(* PLC project HomeAutomation.ecp, WAGO e!COCKPIT e!COCKPIT *)
(* stored: creationDateTime 2022-11-14T18:30:35.868664, modificationDateTime 2022-11-14T18:29:50.9667677 *)

TYPE COVER_STATES : (Idle, Auto, Manual, Prio_up, Prio_dn, Calibrate_up, Calibrate_dn);
END_TYPE

TYPE MQTT_MESSAGE : STRUCT
  Payload : STRING(128);
  Topic : STRING(128);
  Qos : MQTT.QoS;
  MqttRetain : BOOL;
END_STRUCT;
END_TYPE

TYPE RS485_EASTRON_SDM_Devices : (SDM120, SDM220, SDM630);
END_TYPE

TYPE RS485_RtuQuery : STRUCT
  DeviceId : BYTE;
  FunctionCode : BYTE;
  ReadAddress : UINT;
  ReadQuantity : UINT;
END_STRUCT;
END_TYPE

TYPE VIRTUAL_MODES : (Input, Output);
END_TYPE

INTERFACE RS485Device
METHOD RequestBusTime : BOOL
END_METHOD
METHOD GetRtuQuery : RS485_RtuQuery
END_METHOD
METHOD ProcessDataArray
  VAR_INPUT
    Error : POINTER TO BOOL;
    Data : POINTER TO ARRAY[0..124] OF WORD;
  END_VAR
END_METHOD
END_INTERFACE

FUNCTION_BLOCK _RMP_B
  VAR_INPUT
    DIR : BOOL;  (* true = up *)
    E : BOOL := TRUE;
    TR : TIME;
  END_VAR
  VAR_IN_OUT
    RMP : BYTE;
  END_VAR
  VAR
    tx : TIME;
    tl : TIME;
    tn : TIME;
    init : BOOL;
    last_dir : BOOL;
    start : BYTE;
  END_VAR

            (* read system timer *)
tx := DWORD_TO_TIME(OSCAT_BASIC.T_PLC_MS());

IF E AND init AND (dir = last_dir) AND (RMP <> SEL(DIR, 0, 255)) AND TR = tn THEN
	RMP := OSCAT_BASIC.FRMP_B(start, DIR, tx - tl, TR);
ELSE
	init := TRUE;
	tl := tx;
	tn := tr;
	start := RMP;
END_IF;
last_dir := dir;



(* revison history
hm	22. oct. 2008	rev 1.0
	original version

hm	20. nov. 2008	rev 1.1
	set default for E to be TRUE
	added init

hm	19. nov. 2011	rev 1.2
	new code
*)
          

METHOD SetRMP
  VAR_INPUT
    RMP : BYTE;
  END_VAR
                  (*THIS^.RMP:=RMP;*)
THIS^.Start:=RMP;
                
END_METHOD
END_FUNCTION_BLOCK

FUNCTION_BLOCK BLIND_ACTUATOR
  VAR_INPUT
    UP : BOOL;
    DN : BOOL;
    S_IN : BYTE;
    T_UD : TIME := TIME#10s0ms;
    T_ANGLE : TIME := TIME#3s0ms;
    {attribute 'input_constant'}
    T_LOCKOUT : TIME := TIME#100ms;
  END_VAR
  VAR_OUTPUT
    POS : BYTE;
    ANG : BYTE;
    QU : BOOL;
    QD : BOOL;
    STATUS : BYTE;
  END_VAR
  VAR
    position : RMP_B;
    angle : RMP_B;
    lock : OSCAT_BASIC.INTERLOCK;
  END_VAR

            (* make sure only one motor is active at a given time *)
lock(i1 := UP, I2 := DN, TL := T_lockout);

(* ramp up or down to simulate the angle position of the blind slats *)
angle(e := lock.Q1 OR lock.Q2, UP := lock.Q1, PT := T_Angle);
position(e := lock.Q1 AND angle.high OR lock.Q2 AND angle.low, up := lock.Q1, PT := T_UD);

(* set the outputs *)
pos := position.Out;
ang := angle.Out;

(* set the outputs *)
QU := lock.Q1;
QD := lock.Q2;

(* set the status output *)
IF UP AND DN THEN
	 status := 1;			(* error up and down together are not allowed *)
ELSIF UP THEN
	status := 121;
ELSIF DN THEN
	status := 122;
ELSE
	status := S_IN;
END_IF;


(* revision history
hm	29. sep 2007	rev 1.0
	original release

hm	6. oct 2007	rev 1.1
	rearanged outputs

hm	18. oct. 2008	rev 1.2
	changed calls for rmp_B because of change in RMP_B

hm	27. jul. 2009	rev 1.3
	changes status to be 12X

ae	08. mar. 2010 rev 1.4	
	at aPosition

*)
          

METHOD SetPOS
  VAR_INPUT
    POS : BYTE;
  END_VAR
                  THIS^.POS:=POS;
THIS^.position.SetRMP(POS);
                
END_METHOD
END_FUNCTION_BLOCK

FUNCTION CALC_COVER_STATE : COVER_STATES
  VAR_INPUT
    UP : BOOL;
    DN : BOOL;
    PRIO_LOCK : BOOL;
    PRIO_UP : BOOL;
    PRIO_DN : BOOL;
    PI : BYTE;
    POS : BYTE;
    MqttRequestAuto : POINTER TO BOOL;
    MqttRequestStop : POINTER TO BOOL;
    MqttRequestCalibrateUp : POINTER TO BOOL;
    MqttRequestCalibrateDn : POINTER TO BOOL;
    CurrentState : COVER_STATES;
    StateTimer : POINTER TO TOF;
  END_VAR
  VAR
    NewState : COVER_STATES;
  END_VAR

            IF PRIO_LOCK THEN
	NewState := COVER_STATES.Idle;
	MqttRequestAuto^ := FALSE;
	MqttRequestStop^ := FALSE;
	MqttRequestCalibrateUp^ := FALSE;
	MqttRequestCalibrateDn^ := FALSE;
ELSIF PRIO_UP THEN
	NewState := COVER_STATES.Prio_up;
	MqttRequestAuto^ := FALSE;
	MqttRequestStop^ := FALSE;
	MqttRequestCalibrateUp^ := FALSE;
	MqttRequestCalibrateDn^ := FALSE;
ELSIF PRIO_DN THEN
	NewState := COVER_STATES.Prio_dn;
	MqttRequestAuto^ := FALSE;
	MqttRequestStop^ := FALSE;
	MqttRequestCalibrateUp^ := FALSE;
	MqttRequestCalibrateDn^ := FALSE;
ELSIF UP OR DN THEN
	NewState := COVER_STATES.Manual;
	MqttRequestAuto^ := FALSE;
	MqttRequestStop^ := FALSE;
	MqttRequestCalibrateUp^ := FALSE;
	MqttRequestCalibrateDn^ := FALSE;
ELSIF MqttRequestStop^ THEN
	NewState := COVER_STATES.Idle;
	MqttRequestAuto^ := FALSE;
	MqttRequestStop^ := FALSE;
	MqttRequestCalibrateUp^ := FALSE;
	MqttRequestCalibrateDn^ := FALSE;
ELSIF MqttRequestAuto^ AND PI <> POS THEN
	NewState := COVER_STATES.Auto;
	MqttRequestStop^ := FALSE;
	MqttRequestCalibrateUp^ := FALSE;
	MqttRequestCalibrateDn^ := FALSE;
ELSIF MqttRequestAuto^ AND PI = POS THEN
	NewState := COVER_STATES.Idle;
	MqttRequestAuto^ := FALSE;
	MqttRequestStop^ := FALSE;
	MqttRequestCalibrateUp^ := FALSE;
	MqttRequestCalibrateDn^ := FALSE;
ELSIF MqttRequestCalibrateUp^ THEN
	NewState := COVER_STATES.Calibrate_up;
	MqttRequestAuto^ := FALSE;
	MqttRequestStop^ := FALSE;
	MqttRequestCalibrateDn^ := FALSE;
ELSIF MqttRequestCalibrateDn^ THEN
	NewState := COVER_STATES.Calibrate_dn;
	MqttRequestAuto^ := FALSE;
	MqttRequestStop^ := FALSE;
	MqttRequestCalibrateDn^ := FALSE;
ELSE
	NewState := COVER_STATES.Idle;
	MqttRequestAuto^ := FALSE;
	MqttRequestStop^ := FALSE;
	MqttRequestCalibrateUp^ := FALSE;
	MqttRequestCalibrateDn^ := FALSE;
END_IF

IF NewState <> CurrentState THEN
	//Reset StateTimer
	StateTimer^.IN:=TRUE;
END_IF

CALC_COVER_STATE := NewState;
          
END_FUNCTION

{attribute 'reflection'}
FUNCTION_BLOCK FB_INPUT_BINARYSENSOR_MQTT
  VAR_INPUT
    BS : BOOL;
  END_VAR
  VAR_OUTPUT
    Q : BOOL;  (* Follows the input but debounced *)
    EVENT : BOOL;  (* Event outputs only high for on clock cycle *)
    EVENT_R : BOOL;
    EVENT_F : BOOL;
  END_VAR
  VAR
    {attribute 'instance-path'}
    {attribute 'noinit'}
    InstanceName : STRING;  (* object's full instance name *)
    Startup : BOOL := TRUE;
    InitMqttDone : BOOL;
    MqttPublishTopicPrefix : POINTER TO STRING;
    MqttPublishTopicSuffix : STRING(50);
    pMqttPublishQueue : POINTER TO FB_MqttPublishQueue;
    FB_DEBOUNCE : OSCAT_BUILDING.DEBOUNCE;  (* to debounce the physical input *)
    FB_R_TRIG : Standard.R_TRIG;  (* to detect a rising edge on the debounced signal *)
    FB_F_TRIG : Standard.F_TRIG;  (* to detect a falling edge on the debounced signal *)
    T_TurnOffDelay : TIME := TIME#0ms;
    FB_TurnOffDelayTimer : TOF;
  END_VAR

            FB_DEBOUNCE(IN := BS,	
	TD := T#50MS, (* 2x cyle + 10ms *)
	PM := FALSE
	);
	
FB_TurnOffDelayTimer(IN:=FB_DEBOUNCE.Q,
	PT := T_TurnOffDelay,
	Q=>Q
	);

FB_R_TRIG(CLK := FB_TurnOffDelayTimer.Q);
FB_F_TRIG(CLK := FB_TurnOffDelayTimer.Q);

EVENT := FB_R_TRIG.Q OR FB_F_TRIG.Q;
EVENT_R := FB_R_TRIG.Q;
EVENT_F := FB_F_TRIG.Q;

IF (FB_R_TRIG.Q OR (Startup AND FB_DEBOUNCE.Q)) AND InitMqttDone THEN
	pMqttPublishQueue^.AddMessage(
		Payload := 'ON',
		Topic := CONCAT(MqttPublishTopicPrefix^, MqttPublishTopicSuffix),
		Qos := MQTT.QoS.ExactlyOnce,
		MqttRetain := TRUE
	);
	Startup:=FALSE;	
END_IF

IF (FB_F_TRIG.Q OR (Startup AND NOT(FB_DEBOUNCE.Q))) AND InitMqttDone THEN
	pMqttPublishQueue^.AddMessage(
		Payload := 'OFF',
		Topic := CONCAT(MqttPublishTopicPrefix^, MqttPublishTopicSuffix),
		Qos := MQTT.QoS.ExactlyOnce,
		MqttRetain := TRUE
	);
	Startup:=FALSE;	
END_IF
          

METHOD InitMqtt
  VAR_INPUT
    MQTTPublishPrefix : POINTER TO STRING;
    pMqttPublishQueue : POINTER TO FB_MqttPublishQueue;
  END_VAR
  VAR
    InstanceNamePt : POINTER TO STRING;
  END_VAR
                  THIS^.pMqttPublishQueue := pMqttPublishQueue;
THIS^.MqttPublishTopicPrefix := MQTTPublishPrefix;

InstanceNamePt := CommonTypesAndFunctions.FindLastDot(ADR(THIS^.InstanceName)) + 1;
THIS^.MqttPublishTopicSuffix := InstanceNamePt^;

InitMqttDone := TRUE;
                
END_METHOD

METHOD ConfigureFunctionBlock
  VAR_INPUT
    T_TurnOffDelay : TIME;
  END_VAR
                  THIS^.T_TurnOffDelay:=T_TurnOffDelay;
                
END_METHOD
END_FUNCTION_BLOCK

{attribute 'reflection'}
FUNCTION_BLOCK FB_INPUT_PUSHBUTTON_DIMMER_MQTT
  VAR_INPUT
    PB : BOOL;
    SET : BOOL;
    VAL : BYTE;
    RST : BOOL;
  END_VAR
  VAR_OUTPUT
    DIM : BYTE;
    DBL : BOOL;
    Q : BOOL;
    SINGLE : BOOL;
    DOUBLE : BOOL;
    LONG : BOOL;
    P_LONG : BOOL;
  END_VAR
  VAR
    {attribute 'instance-path'}
    {attribute 'noinit'}
    InstanceName : STRING;  (* object's full instance name *)
    InitMqttDone : BOOL;
    MqttPublishTopicPrefix : POINTER TO STRING;
    MqttPublishTopicSuffix : STRING(50);
    pMqttPublishQueue : POINTER TO FB_MqttPublishQueue;
    FB_DIMMER : OSCAT_BUILDING.DIMM_I;
    OutputDimmer : BOOL;
    Qos_Dimm : MQTT.QoS;
    Delta_Dimm : INT;
    FB_DETECTPUSH : OSCAT_BUILDING.CLICK_MODE;
    P_LONG_R_TRIG : Standard.R_TRIG;
    P_LONG_F_TRIG : Standard.F_TRIG;
    PreviousDim : BYTE;  (* Vars to detect statechanges on outputs *)
    PreviousQ : BOOL;
    PreviousDBL : BOOL;
    T_Debounce : TIME := TIME#10ms;  (* Default values for dimmer, can be overwritten by method call *)
    T_Reconfig : TIME := TIME#10s0ms;
    T_On_Max : TIME := TIME#0ms;
    T_Dimm_Start : TIME := TIME#400ms;
    T_Dimm : TIME := TIME#3s0ms;
    Min_On : BYTE := 50;
    Max_On : BYTE := 255;
    Soft_Dimm : BOOL := TRUE;
    Dbl_Toggle : BOOL := FALSE;
    Rst_Out : BOOL := FALSE;
    T_Long : TIME := TIME#400ms;  (* Default value for click mode, can be overwritten by method call *)
  END_VAR

            FB_DIMMER(
	IN:= PB,
	SET:= SET,
	VAL:= VAL,
	RST:= RST,
	OUT:= DIM,
	T_DEBOUNCE:= T_Debounce,
	T_RECONFIG:= T_Reconfig,
	T_ON_MAX:= T_On_Max,
	T_DIMM_START:= T_Dimm_Start,
	T_DIMM:= T_Dimm,
	MIN_ON:= Min_On,
	MAX_ON:= Max_On,
	SOFT_DIMM:= Soft_Dimm,
	DBL_TOGGLE:= Dbl_Toggle,
	RST_OUT:= Rst_Out,
	Q=> Q,
	DBL=> DBL);
	
FB_DETECTPUSH(
	IN:= PB, 	
	SINGLE=> SINGLE, 
	DOUBLE=> DOUBLE, 
	TP_LONG=> LONG, 
	T_LONG:= T_long);
	
P_LONG_R_TRIG(CLK:=FB_DETECTPUSH.LONG);
P_LONG_F_TRIG(CLK:=FB_DETECTPUSH.LONG);
	
IF (ABS(BYTE_TO_INT(PreviousDim) - BYTE_TO_INT(DIM)) >= Delta_Dimm OR PB = FALSE) AND DIM <> PreviousDim AND OutputDimmer AND InitMqttDone  THEN
	PreviousDim:=DIM;
	pMqttPublishQueue^.AddMessage(		
		Payload := BYTE_TO_STRING(DIM),
		Topic := CONCAT(CONCAT(MqttPublishTopicPrefix^, MqttPublishTopicSuffix), '/DIM'),
		Qos := MQTT.QoS.ExactlyOnce,
		MqttRetain := FALSE
	);
END_IF

IF FB_DIMMER.Q <> PreviousQ AND InitMqttDone THEN
	PreviousQ:=FB_DIMMER.Q;
	pMqttPublishQueue^.AddMessage(
		Payload := BOOL_TO_STRING(FB_DIMMER.Q),
		Topic := CONCAT(CONCAT(MqttPublishTopicPrefix^, MqttPublishTopicSuffix), '/Q'),
		Qos := Qos_Dimm,
		MqttRetain := TRUE
	);
END_IF

IF FB_DIMMER.DBL <> PreviousDBL AND InitMqttDone THEN
	PreviousDBL:=FB_DIMMER.DBL;
	pMqttPublishQueue^.AddMessage(
		Payload := BOOL_TO_STRING(FB_DIMMER.DBL),
		Topic := CONCAT(CONCAT(MqttPublishTopicPrefix^, MqttPublishTopicSuffix), '/DBL'),
		Qos := MQTT.QoS.ExactlyOnce,
		MqttRetain := TRUE
	);
END_IF

IF FB_DETECTPUSH.SINGLE AND InitMqttDone THEN
	pMqttPublishQueue^.AddMessage(
		Payload := 'SINGLE',
		Topic := CONCAT(MqttPublishTopicPrefix^, MqttPublishTopicSuffix),
		Qos := MQTT.QoS.ExactlyOnce,
		MqttRetain := FALSE
	);
END_IF

IF FB_DETECTPUSH.DOUBLE AND InitMqttDone THEN
	pMqttPublishQueue^.AddMessage(
		Payload := 'DOUBLE',
		Topic := CONCAT(MqttPublishTopicPrefix^, MqttPublishTopicSuffix),
		Qos := MQTT.QoS.ExactlyOnce,
		MqttRetain := FALSE
	);
END_IF

IF FB_DETECTPUSH.TP_LONG AND InitMqttDone THEN
	pMqttPublishQueue^.AddMessage(
		Payload := 'LONG',
		Topic := CONCAT(MqttPublishTopicPrefix^, MqttPublishTopicSuffix),
		Qos := MQTT.QoS.ExactlyOnce,
		MqttRetain := FALSE
	);
END_IF

IF (P_LONG_R_TRIG.Q OR P_LONG_F_TRIG.Q) AND InitMqttDone THEN
	pMqttPublishQueue^.AddMessage(
		Payload := BOOL_TO_STRING(FB_DETECTPUSH.LONG),
		Topic := CONCAT(CONCAT(MqttPublishTopicPrefix^, MqttPublishTopicSuffix),'/P_LONG'),
		Qos := MQTT.QoS.ExactlyOnce,
		MqttRetain := TRUE
	);
END_IF
          

METHOD InitMqtt
  VAR_INPUT
    MQTTPublishPrefix : POINTER TO STRING;
    pMqttPublishQueue : POINTER TO FB_MqttPublishQueue;
    OutputDimmer : BOOL;
    Qos_Dimm : MQTT.QoS;
    Delta_Dimm : INT;
  END_VAR
  VAR
    InstanceNamePt : POINTER TO STRING;
  END_VAR
                  THIS^.pMqttPublishQueue := pMqttPublishQueue;
THIS^.MqttPublishTopicPrefix := MQTTPublishPrefix;

InstanceNamePt := CommonTypesAndFunctions.FindLastDot(ADR(THIS^.InstanceName)) + 1;
THIS^.MqttPublishTopicSuffix := InstanceNamePt^;

THIS^.OutputDimmer:=OutputDimmer;
THIS^.Qos_Dimm:=Qos_Dimm;
THIS^.Delta_Dimm:=Delta_Dimm;

InitMqttDone := TRUE;
                
END_METHOD

METHOD ConfigureFunctionBlock
  VAR_INPUT
    T_Debounce : TIME;  (* Default values for dimmer, can be overwritten by method call *)
    T_Reconfig : TIME;
    T_On_Max : TIME;
    T_Dimm_Start : TIME;
    T_Dimm : TIME;
    Min_On : BYTE;
    Max_On : BYTE;
    Soft_Dimm : BOOL;
    Dbl_Toggle : BOOL;
    Rst_Out : BOOL;
    T_Long : TIME;  (* Default value for click mode, can be overwritten by method call *)
  END_VAR
                  THIS^.T_Debounce:=T_Debounce;
THIS^.T_Reconfig:=T_Reconfig;
THIS^.T_On_Max:=T_On_Max;
THIS^.T_Dimm_Start:=T_Dimm_Start;
THIS^.T_Dimm:=T_Dimm;
THIS^.Min_On:=Min_On;
THIS^.Max_On:=Max_On;

THIS^.T_Long:=T_Long;
                
END_METHOD
END_FUNCTION_BLOCK

{attribute 'reflection'}
FUNCTION_BLOCK FB_INPUT_PUSHBUTTON_MQTT
  VAR_INPUT
    PB : BOOL;
  END_VAR
  VAR_OUTPUT
    SINGLE : BOOL;
    DOUBLE : BOOL;
    LONG : BOOL;
    P_LONG : BOOL;
  END_VAR
  VAR
    {attribute 'instance-path'}
    {attribute 'noinit'}
    InstanceName : STRING;  (* object's full instance name *)
    InitMqttDone : BOOL;
    MqttPublishTopicPrefix : POINTER TO STRING;
    MqttPublishTopicSuffix : STRING(50);
    pMqttPublishQueue : POINTER TO FB_MqttPublishQueue;
    FB_DETECTPUSH : OSCAT_BUILDING.CLICK_MODE;
    P_LONG_R_TRIG : Standard.R_TRIG;
    P_LONG_F_TRIG : Standard.F_TRIG;
    T_Long : TIME := TIME#400ms;  (* Default value for click mode, can be overwritten by method call *)
  END_VAR

            FB_DETECTPUSH(
	IN:= PB, 	
	SINGLE=> SINGLE, 
	DOUBLE=> DOUBLE, 
	TP_LONG=> LONG, 
	LONG=> P_LONG,
	T_LONG:= T_Long);
	
P_LONG_R_TRIG(CLK:=FB_DETECTPUSH.LONG);
P_LONG_F_TRIG(CLK:=FB_DETECTPUSH.LONG);
	
IF FB_DETECTPUSH.SINGLE AND InitMqttDone THEN
	pMqttPublishQueue^.AddMessage(
		Payload := 'SINGLE',
		Topic := CONCAT(MqttPublishTopicPrefix^, MqttPublishTopicSuffix),
		Qos := MQTT.QoS.ExactlyOnce,
		MqttRetain := FALSE
	);
END_IF

IF FB_DETECTPUSH.DOUBLE AND InitMqttDone THEN
	pMqttPublishQueue^.AddMessage(
		Payload := 'DOUBLE',
		Topic := CONCAT(MqttPublishTopicPrefix^, MqttPublishTopicSuffix),
		Qos := MQTT.QoS.ExactlyOnce,
		MqttRetain := FALSE
	);
END_IF

IF FB_DETECTPUSH.TP_LONG AND InitMqttDone THEN
	pMqttPublishQueue^.AddMessage(
		Payload := 'LONG',
		Topic := CONCAT(MqttPublishTopicPrefix^, MqttPublishTopicSuffix),
		Qos := MQTT.QoS.ExactlyOnce,
		MqttRetain := FALSE
	);
END_IF

IF (P_LONG_R_TRIG.Q OR P_LONG_F_TRIG.Q) AND InitMqttDone THEN
	pMqttPublishQueue^.AddMessage(
		Payload := BOOL_TO_STRING(FB_DETECTPUSH.LONG),
		Topic := CONCAT(CONCAT(MqttPublishTopicPrefix^, MqttPublishTopicSuffix),'/P_LONG'),
		Qos := MQTT.QoS.ExactlyOnce,
		MqttRetain := TRUE
	);
END_IF
          

METHOD InitMqtt
  VAR_INPUT
    MQTTPublishPrefix : POINTER TO STRING;
    pMqttPublishQueue : POINTER TO FB_MqttPublishQueue;
  END_VAR
  VAR
    InstanceNamePt : POINTER TO STRING;
  END_VAR
                  THIS^.pMqttPublishQueue := pMqttPublishQueue;
THIS^.MqttPublishTopicPrefix := MQTTPublishPrefix;

InstanceNamePt := CommonTypesAndFunctions.FindLastDot(ADR(THIS^.InstanceName)) + 1;
THIS^.MqttPublishTopicSuffix := InstanceNamePt^;

InitMqttDone := TRUE;
                
END_METHOD

METHOD ConfigureFunctionBlock
  VAR_INPUT
    T_Long : TIME;  (* Default value for click mode, can be overwritten by method call *)
  END_VAR
                  THIS^.T_Long:=T_Long;
                
END_METHOD
END_FUNCTION_BLOCK

FUNCTION_BLOCK FB_MqttPublishQueue
  VAR_OUTPUT
    EMPTY : BOOL := TRUE;
    FULL : BOOL;
  END_VAR
  VAR
    localMessage : MQTT_MESSAGE;
    fifo : ARRAY[0..n] OF MQTT_MESSAGE;
    pr : INT;
    pw : INT;
  END_VAR
  VAR CONSTANT
    n : INT := 1024;  (* changing this value will chage the number of stored elements in the fifo *)
  END_VAR

            
          

METHOD GetMessage : MQTT_MESSAGE
                  IF NOT EMPTY THEN
	GetMessage := fifo[pr];
	pr := OSCAT_BASIC.INC1(pr,n);
	EMPTY := pr = pw;
	FULL := FALSE;
END_IF;
                
END_METHOD

METHOD AddMessage
  VAR_INPUT
    Payload : STRING(128);
    Topic : STRING(128);
    Qos : MQTT.QoS;
    MqttRetain : BOOL;
  END_VAR
                  IF NOT FULL THEN
	localMessage.Payload := Payload;
	localMessage.Topic := Topic;
	localMessage.Qos := Qos;
	localMessage.MqttRetain := MqttRetain;
	fifo[pw] := localMessage;
	pw := OSCAT_BASIC.INC1(pw,n);
	FULL := pw = pr;
	EMPTY := FALSE;
END_IF;
                
END_METHOD

METHOD Reset
                  pw := pr;
FULL := FALSE;
EMPTY := TRUE;
                
END_METHOD
END_FUNCTION_BLOCK

FUNCTION_BLOCK FB_MqttPublishWorker
  VAR_OUTPUT
    SendDone : BOOL;
  END_VAR
  VAR
    LocalMqttMessage : MQTT_MESSAGE;
    InitDone : BOOL;
    RequestToSend : BOOL;
    Send : BOOL;
    publish : MQTT.MQTTPublish;
  END_VAR

            //need to call publish here because of FB nums
publish(
	Topic:= ADR(LocalMqttMessage.Topic), 
	PayloadString:= ADR(LocalMqttMessage.Payload), 
	PublishAsString:= TRUE, 
	QoSIn:= LocalMqttMessage.Qos, 
	MRetain:= LocalMqttMessage.MqttRetain, 
	send:= Send);
	
IF NOT InitDone THEN RETURN; END_IF

IF RequestToSend THEN
	Send := TRUE;
	SendDone := FALSE;
END_IF

IF publish.done THEN
	 SendDone := TRUE;
	 RequestToSend:=FALSE;
	 Send:=FALSE;
END_IF
          

METHOD Init
  VAR_INPUT
    inputMQTT_IN_OUT : POINTER TO MQTT.MQTT_IN_OUT;  (* Pointer MQTTT exchange strucure *)
  END_VAR
                  publish.SetMqttInOut(MQTT_IN_OUT := inputMQTT_IN_OUT^);

InitDone := TRUE;
SendDone := TRUE;

                
END_METHOD

METHOD PublishMessage
  VAR_INPUT
    MqttMessage : MQTT_MESSAGE;
  END_VAR
                  LocalMqttMessage := MqttMessage;

RequestToSend:=TRUE;
                
END_METHOD
END_FUNCTION_BLOCK

{attribute 'reflection'}
FUNCTION_BLOCK FB_OUTPUT_BISTABLE_MQTT IMPLEMENTS MQTT.MQTT_SUBSCRIBE_CALLBACK
  VAR_INPUT
    PRIO_HIGH : BOOL := FALSE;
    PRIO_LOW : BOOL := FALSE;
    TOGGLE : BOOL := FALSE;
    FEEDBACK : BOOL := FALSE;
  END_VAR
  VAR_OUTPUT
    OUT : BOOL;
  END_VAR
  VAR
    {attribute 'instance-path'}
    {attribute 'noinit'}
    InstanceName : STRING;  (* object's full instance name *)
    Startup : BOOL := TRUE;
    InitMqttDone : BOOL;
    MqttPublishTopicPrefix : POINTER TO STRING;
    MqttPublishTopicSuffix : STRING(50);
    MQTTSubscribeTopic : STRING(50);
    pMqttPublishQueue : POINTER TO FB_MqttPublishQueue;
    MqttHighRequest : BOOL;
    MqttLowRequest : BOOL;
    PreviousFeedback : BOOL;
    HoldTimer : TOF;
    T_hold : TIME := TIME#1s0ms;
    PulseTrigger : BOOL := FALSE;
  END_VAR

            HoldTimer(PT:= T_hold);

IF PRIO_HIGH THEN
	IF NOT FEEDBACK THEN
		PulseTrigger:=TRUE;
	END_IF
ELSIF(PRIO_LOW AND NOT (PRIO_HIGH)) THEN
	IF FEEDBACK THEN		
		PulseTrigger:=TRUE;
	END_IF
	OUT:= FALSE;
ELSIF MqttHighRequest THEN
	IF NOT FEEDBACK THEN		
		PulseTrigger:=TRUE;
	END_IF
	MqttHighRequest := FALSE;
	MqttLowRequest := FALSE;
ELSIF MqttLowRequest THEN
	IF FEEDBACK THEN		
		PulseTrigger:=TRUE;
	END_IF
	MqttHighRequest := FALSE;
	MqttLowRequest := FALSE;
ELSIF(TOGGLE) THEN	
	PulseTrigger:=TRUE;
END_IF;

IF ((PreviousFeedback <> FEEDBACK) OR Startup) AND InitMqttDone THEN
	pMqttPublishQueue^.AddMessage(
		Payload := BOOL_TO_STRING(FEEDBACK),
		Topic := CONCAT(MqttPublishTopicPrefix^, MqttPublishTopicSuffix),
		Qos := MQTT.QoS.ExactlyOnce,
		MqttRetain := TRUE
	);	
	Startup:=FALSE;
END_IF	

PreviousFeedback := FEEDBACK;
HoldTimer.IN	 := PulseTrigger;
OUT := HoldTimer.Q;

PulseTrigger:=FALSE;
          

METHOD InitMqtt
  VAR_INPUT
    MQTTPublishPrefix : POINTER TO STRING;
    MQTTSubscribePrefix : POINTER TO STRING;
    pMqttPublishQueue : POINTER TO FB_MqttPublishQueue;
    pMqttCallbackCollector : POINTER TO MQTT.CallbackCollector;
  END_VAR
  VAR
    InstanceNamePt : POINTER TO STRING;
  END_VAR
                  THIS^.pMqttPublishQueue := pMqttPublishQueue;
THIS^.MqttPublishTopicPrefix := MQTTPublishPrefix;

InstanceNamePt := CommonTypesAndFunctions.FindLastDot(ADR(THIS^.InstanceName)) + 1;
THIS^.MqttPublishTopicSuffix := InstanceNamePt^;
THIS^.MQTTSubscribeTopic := CONCAT(MQTTSubscribePrefix^ ,THIS^.MqttPublishTopicSuffix);

// register the FB agains the collector so mqtt events can be received
pMqttCallbackCollector^.put(instance:= THIS^);

InitMqttDone := TRUE;
                
END_METHOD

METHOD PublishReceived : BOOL
  VAR_INPUT
    Data : MQTT.CALLBACK_DATA;  (* Collection of recived Data *)
  END_VAR
                  //first check if Mqtt is initialized, otherwise do nothing
IF NOT(InitMqttDone) THEN
	//mark the interface call from the collector as done
	PublishReceived := TRUE;
//check if the packet is for this FB
ELSIF CommonTypesAndFunctions.StrEquals(str1:= ADR(MQTTSubscribeTopic), str2:= Data.TopicOut) THEN
	//mark the interface call from the collector as done
	PublishReceived := TRUE;
	//now process the data
	IF CommonTypesAndFunctions.StrEquals(str1:= Data.PayloadString, str2:= ADR('TRUE')) THEN
		MqttHighRequest := TRUE;
	END_IF
	IF CommonTypesAndFunctions.StrEquals(str1:= Data.PayloadString, str2:= ADR('FALSE')) THEN
		MqttLowRequest := TRUE;
	END_IF
END_IF 
                
END_METHOD

METHOD ConfigureFunctionBlock
  VAR_INPUT
    T_hold : TIME;  (* Default value for click mode, can be overwritten by method call *)
  END_VAR
                  THIS^.T_hold:=T_hold;
                
END_METHOD
END_FUNCTION_BLOCK

{attribute 'reflection'}
FUNCTION_BLOCK FB_OUTPUT_COVER_MQTT IMPLEMENTS MQTT.MQTT_SUBSCRIBE_CALLBACK
  VAR_INPUT
    UP : BOOL;
    DN : BOOL;
    PI : BYTE;
    PRIO_LOCK : BOOL;
    PRIO_UP : BOOL;
    PRIO_DN : BOOL;
    {attribute 'input_constant'}
    SENS : BYTE := 1;
    {attribute 'input_constant'}
    T_LOCKOUT : TIME := TIME#1s0ms;
    {attribute 'input_constant'}
    T_UD : TIME := TIME#10s0ms;
  END_VAR
  VAR_OUTPUT
    POS : BYTE;
    MU : BOOL;
    MD : BOOL;
  END_VAR
  VAR
    {attribute 'instance-path'}
    {attribute 'noinit'}
    InstanceName : STRING;  (* object's full instance name *)
    Startup : BOOL := TRUE;
    InitMqttDone : BOOL;
    MqttPublishTopicPrefix : POINTER TO STRING;
    MqttPublishTopicSuffix : STRING(50);
    MQTTSubscribeTopic : STRING(50);
    pMqttPublishQueue : POINTER TO FB_MqttPublishQueue;
    FB_ACT : BLIND_ACTUATOR;
    delta : BYTE;
    internal_UP : BOOL;
    internal_DN : BOOL;
    Qos_POS : MQTT.QoS;
    Delta_POS : INT;
    Cover_State : COVER_STATES;
    Cover_State_Timer : TOF;
    MqttRequestAuto : BOOL;
    MqttRequestStop : BOOL;
    MqttRequestCalibrateUp : BOOL;
    MqttRequestCalibrateDn : BOOL;
  END_VAR
  VAR PERSISTENT
    PreviousPos : BYTE;  (* To retain position through powercycles *)
  END_VAR

            IF Startup THEN
	POS:=PreviousPos;
	FB_ACT.SetPOS(PreviousPos);
END_IF

Cover_State_Timer(PT:=2 * T_UD);
Cover_State_Timer.IN:=FALSE;

CASE Cover_State OF
	COVER_STATES.Idle:
		internal_UP:=FALSE;
		internal_DN:=FALSE;
		//Calculate the next state
		Cover_State := CALC_COVER_STATE(UP:=UP,DN:=DN,PRIO_LOCK:=PRIO_LOCK,PRIO_UP:=PRIO_UP,PRIO_DN:=PRIO_DN,PI:=PI,POS:=POS,MqttRequestAuto:=ADR(MqttRequestAuto),MqttRequestStop:=ADR(MqttRequestStop),MqttRequestCalibrateUp:=ADR(MqttRequestCalibrateUp),MqttRequestCalibrateDn:=ADR(MqttRequestCalibrateDn),CurrentState:=Cover_State,StateTimer:=ADR(Cover_State_Timer));
	COVER_STATES.Prio_up:
		// Only power an engine for maximum twice T_UD
		IF Cover_State_Timer.Q THEN
			internal_UP:=TRUE;
			internal_DN:=FALSE;
		ELSE
			internal_UP:=FALSE;
			internal_DN:=FALSE;
		END_IF
		//Calculate the next state
		Cover_State := CALC_COVER_STATE(UP:=UP,DN:=DN,PRIO_LOCK:=PRIO_LOCK,PRIO_UP:=PRIO_UP,PRIO_DN:=PRIO_DN,PI:=PI,POS:=POS,MqttRequestAuto:=ADR(MqttRequestAuto),MqttRequestStop:=ADR(MqttRequestStop),MqttRequestCalibrateUp:=ADR(MqttRequestCalibrateUp),MqttRequestCalibrateDn:=ADR(MqttRequestCalibrateDn),CurrentState:=Cover_State,StateTimer:=ADR(Cover_State_Timer));
	COVER_STATES.Prio_dn:
		// Only power an engine for maximum twice T_UD
		IF Cover_State_Timer.Q THEN
			internal_UP:=FALSE;
			internal_DN:=TRUE;
		ELSE
			internal_UP:=FALSE;
			internal_DN:=FALSE;
		END_IF
		//Calculate the next state
		Cover_State := CALC_COVER_STATE(UP:=UP,DN:=DN,PRIO_LOCK:=PRIO_LOCK,PRIO_UP:=PRIO_UP,PRIO_DN:=PRIO_DN,PI:=PI,POS:=POS,MqttRequestAuto:=ADR(MqttRequestAuto),MqttRequestStop:=ADR(MqttRequestStop),MqttRequestCalibrateUp:=ADR(MqttRequestCalibrateUp),MqttRequestCalibrateDn:=ADR(MqttRequestCalibrateDn),CurrentState:=Cover_State,StateTimer:=ADR(Cover_State_Timer));
	COVER_STATES.Auto:
		internal_UP:=TRUE;
		internal_DN:=TRUE;
		//Calculate the next state
		Cover_State := CALC_COVER_STATE(UP:=UP,DN:=DN,PRIO_LOCK:=PRIO_LOCK,PRIO_UP:=PRIO_UP,PRIO_DN:=PRIO_DN,PI:=PI,POS:=POS,MqttRequestAuto:=ADR(MqttRequestAuto),MqttRequestStop:=ADR(MqttRequestStop),MqttRequestCalibrateUp:=ADR(MqttRequestCalibrateUp),MqttRequestCalibrateDn:=ADR(MqttRequestCalibrateDn),CurrentState:=Cover_State,StateTimer:=ADR(Cover_State_Timer));
	COVER_STATES.Manual:
		internal_UP:=UP;
		internal_DN:=DN;
		//Calculate the next state
		Cover_State := CALC_COVER_STATE(UP:=UP,DN:=DN,PRIO_LOCK:=PRIO_LOCK,PRIO_UP:=PRIO_UP,PRIO_DN:=PRIO_DN,PI:=PI,POS:=POS,MqttRequestAuto:=ADR(MqttRequestAuto),MqttRequestStop:=ADR(MqttRequestStop),MqttRequestCalibrateUp:=ADR(MqttRequestCalibrateUp),MqttRequestCalibrateDn:=ADR(MqttRequestCalibrateDn),CurrentState:=Cover_State,StateTimer:=ADR(Cover_State_Timer));
	COVER_STATES.Calibrate_up:
		// Only power an engine for maximum twice T_UD
		IF Cover_State_Timer.Q THEN
			internal_UP:=FALSE;
			internal_DN:=TRUE;
		ELSE
			internal_UP:=FALSE;
			internal_DN:=FALSE;
			//Finish the request
			MqttRequestCalibrateUp:=FALSE;
		END_IF
		//Calculate the next state
		Cover_State := CALC_COVER_STATE(UP:=UP,DN:=DN,PRIO_LOCK:=PRIO_LOCK,PRIO_UP:=PRIO_UP,PRIO_DN:=PRIO_DN,PI:=PI,POS:=POS,MqttRequestAuto:=ADR(MqttRequestAuto),MqttRequestStop:=ADR(MqttRequestStop),MqttRequestCalibrateUp:=ADR(MqttRequestCalibrateUp),MqttRequestCalibrateDn:=ADR(MqttRequestCalibrateDn),CurrentState:=Cover_State,StateTimer:=ADR(Cover_State_Timer));
	COVER_STATES.Calibrate_dn:
		// Only power an engine for maximum twice T_UD
		IF Cover_State_Timer.Q THEN
			internal_UP:=FALSE;
			internal_DN:=TRUE;
		ELSE
			internal_UP:=FALSE;
			internal_DN:=FALSE;
			//Finish the request
			MqttRequestCalibrateDn:=FALSE;
		END_IF
		//Calculate the next state
		Cover_State := CALC_COVER_STATE(UP:=UP,DN:=DN,PRIO_LOCK:=PRIO_LOCK,PRIO_UP:=PRIO_UP,PRIO_DN:=PRIO_DN,PI:=PI,POS:=POS,MqttRequestAuto:=ADR(MqttRequestAuto),MqttRequestStop:=ADR(MqttRequestStop),MqttRequestCalibrateUp:=ADR(MqttRequestCalibrateUp),MqttRequestCalibrateDn:=ADR(MqttRequestCalibrateDn),CurrentState:=Cover_State,StateTimer:=ADR(Cover_State_Timer));
	ELSE
		Cover_State:=COVER_STATES.Idle;
END_CASE

(* Check Position*)
FB_ACT(T_UD:=T_UD, T_ANGLE:=T#0S, T_lockout := T_Lockout);

IF internal_UP AND internal_DN THEN
	(* automatic modus detected *)
	(* first find correct position *)
	IF BYTE_TO_INT(FB_ACT.pos) < BYTE_TO_INT(pi) - delta THEN
		FB_ACT.UP := TRUE;
		FB_ACT.DN := FALSE;
		delta := 0;
	ELSIF BYTE_TO_INT(FB_ACT.pos) > BYTE_TO_INT(pi) + delta THEN
		FB_ACT.UP := FALSE;
		FB_ACT.DN := TRUE;
		delta := 0;
	(* correct position reached *)
	ELSE
		FB_ACT.UP := FALSE;
		FB_ACT.DN := FALSE;
		delta := sens;
	END_IF;
ELSE
	FB_ACT.UP := internal_UP;
	FB_ACT.DN := internal_DN;
END_IF;

(* blind control calls blind_actuator *)
FB_ACT(T_UD:=T_UD, T_ANGLE:=T#0S, T_lockout := T_Lockout);
POS := FB_ACT.pos;
MU := FB_ACT.QU;
MD := FB_ACT.QD;

IF ((ABS(BYTE_TO_INT(PreviousPos) - BYTE_TO_INT(POS)) >= Delta_POS  OR (MU = FALSE AND MD = FALSE)) AND POS <> PreviousPos OR Startup) AND InitMqttDone THEN
	PreviousPos:=POS;
	pMqttPublishQueue^.AddMessage(
		Payload := INT_TO_STRING(REAL_TO_INT(OSCAT_BASIC.SCALE_B(X:=POS, I_LO:=0, I_HI:=255, O_LO:=0, O_HI:=100))),
		Topic := CONCAT(MqttPublishTopicPrefix^, MqttPublishTopicSuffix),
		Qos := Qos_POS,
		MqttRetain := TRUE
	);
	Startup:=FALSE;
END_IF

          

METHOD InitMqtt
  VAR_INPUT
    MQTTPublishPrefix : POINTER TO STRING;
    MQTTSubscribePrefix : POINTER TO STRING;
    pMqttPublishQueue : POINTER TO FB_MqttPublishQueue;
    pMqttCallbackCollector : POINTER TO MQTT.CallbackCollector;
    Qos_POS : MQTT.QoS;
    Delta_POS : INT;
  END_VAR
  VAR
    InstanceNamePt : POINTER TO STRING;
  END_VAR
                  THIS^.pMqttPublishQueue := pMqttPublishQueue;
THIS^.MqttPublishTopicPrefix := MQTTPublishPrefix;

InstanceNamePt := CommonTypesAndFunctions.FindLastDot(ADR(THIS^.InstanceName)) + 1;
THIS^.MqttPublishTopicSuffix := InstanceNamePt^;
THIS^.MQTTSubscribeTopic := CONCAT(MQTTSubscribePrefix^ ,THIS^.MqttPublishTopicSuffix);

// register the FB agains the collector so mqtt events can be received
pMqttCallbackCollector^.put(instance:= THIS^);

THIS^.Qos_POS:=Qos_POS;
THIS^.Delta_POS:=REAL_TO_INT(OSCAT_BASIC.SCALE_B(X:=INT_TO_BYTE(Delta_POS), I_LO:=0, I_HI:=100, O_LO:=0, O_HI:=255));

InitMqttDone := TRUE;
                
END_METHOD

METHOD PublishReceived : BOOL
  VAR_INPUT
    Data : MQTT.CALLBACK_DATA;  (* Collection of recived Data *)
  END_VAR
                  //first check if Mqtt is initialized, otherwise do nothing
IF NOT(InitMqttDone) THEN
	//mark the interface call from the collector as done
	PublishReceived := TRUE;
//check if the packet is for this FB
ELSIF CommonTypesAndFunctions.StrEquals(str1:= ADR(MQTTSubscribeTopic), str2:= Data.TopicOut) THEN
	//mark the interface call from the collector as done
	PublishReceived := TRUE;
	//now process the data
	IF CommonTypesAndFunctions.StrEquals(str1:= Data.PayloadString, str2:= ADR('STOP')) THEN			
		THIS^.MqttRequestStop:=TRUE;
	ELSIF CommonTypesAndFunctions.StrEquals(str1:= Data.PayloadString, str2:= ADR('OPEN')) THEN
		THIS^.PI:=255;
		THIS^.MqttRequestAuto:=TRUE;
	ELSIF CommonTypesAndFunctions.StrEquals(str1:= Data.PayloadString, str2:= ADR('CLOSE')) THEN		
		THIS^.PI:=0;
		THIS^.MqttRequestAuto:=TRUE;
	ELSIF CommonTypesAndFunctions.StrEquals(str1:= Data.PayloadString, str2:= ADR('CAL_UP')) THEN
		THIS^.MqttRequestCalibrateUp:=TRUE;
	ELSIF CommonTypesAndFunctions.StrEquals(str1:= Data.PayloadString, str2:= ADR('CAL_DN')) THEN
		THIS^.MqttRequestCalibrateDn:=TRUE;
	ELSIF OSCAT_BASIC.IS_NUM(str:= Data.PayloadString^) THEN
		THIS^.PI:=REAL_TO_BYTE(OSCAT_BASIC.SCALE_B(X:=STRING_TO_BYTE(Data.PayloadString^), I_LO:=0, I_HI:=100, O_LO:=0, O_HI:=255));
		THIS^.MqttRequestAuto:=TRUE;
	END_IF

END_IF 
                
END_METHOD

METHOD ConfigureFunctionBlock : BOOL
  VAR_INPUT
    T_LOCKOUT : TIME;
    T_UD : TIME;
  END_VAR
                  THIS^.T_LOCKOUT:=T_LOCKOUT;
THIS^.T_UD:=T_UD;
                
END_METHOD
END_FUNCTION_BLOCK

{attribute 'reflection'}
FUNCTION_BLOCK FB_OUTPUT_DIMMER_MQTT IMPLEMENTS MQTT.MQTT_SUBSCRIBE_CALLBACK
  VAR_INPUT
    SINGLE : BOOL;
    LONG : BOOL;
    P_LONG : BOOL;
    PRIO_HIGH : BOOL := FALSE;
    PRIO_LOW : BOOL := FALSE;
    SET : BOOL;
    VAL : BYTE;
    RST : BOOL;
  END_VAR
  VAR_OUTPUT
    Q : BOOL;
    Q_OUT : WORD;
    OUT : WORD;
  END_VAR
  VAR
    t3 : OSCAT_BASIC.TON;
    dim : OSCAT_BASIC._RMP_B;
    dir : BOOL;
    OUT_Internal : BYTE;
    LIN_TRAFO : Util.LIN_TRAFO;
    OUT_LinearScaleMin : INT := 0;
    OUT_LinearScaleMax : INT := 32767;
    {attribute 'instance-path'}
    {attribute 'noinit'}
    InstanceName : STRING;  (* object's full instance name *)
    Startup : BOOL := TRUE;
    InitMqttDone : BOOL;
    MqttPublishTopicPrefix : POINTER TO STRING;
    MqttPublishTopicSuffix : STRING(50);
    MQTTSubscribeTopic : STRING(50);
    pMqttPublishQueue : POINTER TO FB_MqttPublishQueue;
    OutputDimmer : BOOL;
    Qos_Dimm : MQTT.QoS;
    Delta_Dimm : INT;
    T_Debounce : TIME := TIME#10ms;  (* Default values for dimmer, can be overwritten by method call *)
    T_Reconfig : TIME := TIME#10s0ms;
    T_On_Max : TIME := TIME#0ms;
    T_Dimm_Start : TIME := TIME#400ms;
    T_Dimm : TIME := TIME#3s0ms;
    Min_On : BYTE := 50;
    Max_On : BYTE := 255;
    Soft_Dimm : BOOL := TRUE;
    Rst_Out : BOOL := FALSE;
    MqttHighRequest : BOOL;
    MqttLowRequest : BOOL;
  END_VAR
  VAR PERSISTENT
    PreviousOUT : BYTE;  (* To retain output state through powercycles *)
    PreviousQ : BOOL;  (* To retain output state through powercycles *)
  END_VAR

            IF Startup THEN
	OUT := PreviousOUT;
	Q := PreviousQ;
END_IF

IF RST THEN
	IF rst_out THEN OUT_Internal := 0; END_IF;
	Q := FALSE;
	dir := OUT_Internal > 127;
ELSIF PRIO_HIGH THEN
	Q := TRUE;
	OUT_Internal := 255;
ELSIF PRIO_LOW THEN
	Q := FALSE;
ELSIF MqttHighRequest THEN
	Q:= TRUE;
	MqttHighRequest := FALSE;
	MqttLowRequest := FALSE;
ELSIF MqttLowRequest THEN
	Q:= FALSE;
	MqttHighRequest := FALSE;
	MqttLowRequest := FALSE;
ELSIF set THEN
	OUT_Internal := val;
	Q := TRUE;
	(* set direction to up when value < 127 otherwise set dir down dir is reversed because next action will reverse again *)
	dir := OUT_Internal > 127;
ELSIF SINGLE THEN
	(* a single click reverses output Q *)
	Q := NOT Q;
	(* when dimmer is turned on we need to limit out to min and max limits *)
	IF Q THEN OUT_Internal := LIMIT(MAX(OUT_Internal,1), OUT_Internal, MAX_ON);	END_IF;
	(* set the appropriate direction of dimmer dir is reversed because next action will reverse again *)
	dir := OUT_Internal > 127;
ELSIF LONG THEN
	IF NOT Q THEN
		IF SOFT_DIMM THEN
			OUT_Internal := 1;
			dir := TRUE;
		ELSE
			OUT_Internal := LIMIT(MAX(MIN_ON,1), OUT_Internal, MAX_ON);
			DIR := OUT_Internal < 127;
		END_IF;
		Q := TRUE;
	ELSE
		(* reverse direction with every long click *)
		dir := NOT dir;
	END_IF;
END_IF;


(* while dimming is active ramp the output out up or down *)
dim(DIR := dir, e := P_LONG AND Q, TR := T_DIMM, rmp := OUT_Internal);

(* reverse direction when limits are reached *)
IF OUT_Internal = 0 THEN
	dir := TRUE;
ELSIF OUT_Internal = 255 THEN
	dir := FALSE;
END_IF;

(* limit the maximum runtime *)
IF t_ON_MAX > t#0s THEN
	t3(in := q, pt := T_ON_MAX);
	Q := Q XOR t3.Q;
END_IF;

(* Scale the internal OUT to the actual OUT *)
LIN_TRAFO(
		IN:= OUT_Internal,
		IN_MIN:= 0,
		IN_MAX:= 255,
		OUT_MIN:=OUT_LinearScaleMin,
		OUT_MAX:=OUT_LinearScaleMax
	);
OUT:= REAL_TO_WORD(LIN_TRAFO.OUT);
IF Q THEN
	Q_OUT:= OUT;
ELSE
	Q_OUT:= 0;
END_IF

IF ((ABS(BYTE_TO_INT(PreviousOUT) - BYTE_TO_INT(OUT_Internal)) >= Delta_Dimm) OR Startup AND OUT_Internal <> PreviousOUT OR Startup AND OutputDimmer) AND InitMqttDone THEN
	PreviousOUT:=OUT_Internal;
	pMqttPublishQueue^.AddMessage(		
		Payload := BYTE_TO_STRING(OUT_Internal),
		Topic := CONCAT(CONCAT(MqttPublishTopicPrefix^, MqttPublishTopicSuffix), '/OUT'),
		Qos := MQTT.QoS.ExactlyOnce,
		MqttRetain := TRUE
	);
END_IF

IF (Q <> PreviousQ OR Startup) AND InitMqttDone THEN
	PreviousQ:=Q;
	pMqttPublishQueue^.AddMessage(
		Payload := BOOL_TO_STRING(Q),
		Topic := CONCAT(CONCAT(MqttPublishTopicPrefix^, MqttPublishTopicSuffix), '/Q'),
		Qos := Qos_Dimm,
		MqttRetain := TRUE
	);
END_IF

Startup:=FALSE;


          

METHOD InitMqtt
  VAR_INPUT
    MQTTPublishPrefix : POINTER TO STRING;
    MQTTSubscribePrefix : POINTER TO STRING;
    pMqttPublishQueue : POINTER TO FB_MqttPublishQueue;
    pMqttCallbackCollector : POINTER TO MQTT.CallbackCollector;
    OutputDimmer : BOOL;
    Qos_Dimm : MQTT.QoS;
    Delta_Dimm : INT;
  END_VAR
  VAR
    InstanceNamePt : POINTER TO STRING;
  END_VAR
                  THIS^.pMqttPublishQueue := pMqttPublishQueue;
THIS^.MqttPublishTopicPrefix := MQTTPublishPrefix;

InstanceNamePt := CommonTypesAndFunctions.FindLastDot(ADR(THIS^.InstanceName)) + 1;
THIS^.MqttPublishTopicSuffix := InstanceNamePt^;
THIS^.MQTTSubscribeTopic := CONCAT(MQTTSubscribePrefix^ ,THIS^.MqttPublishTopicSuffix);

THIS^.OutputDimmer:=OutputDimmer;
THIS^.Qos_Dimm:=Qos_Dimm;
THIS^.Delta_Dimm:=Delta_Dimm;

// register the FB agains the collector so mqtt events can be received
pMqttCallbackCollector^.put(instance:= THIS^);

InitMqttDone := TRUE;
                
END_METHOD

METHOD ConfigureFunctionBlock
  VAR_INPUT
    T_Debounce : TIME;  (* Default values for dimmer, can be overwritten by method call *)
    T_Reconfig : TIME;
    T_On_Max : TIME;
    T_Dimm_Start : TIME;
    T_Dimm : TIME;
    Min_On : BYTE;
    Max_On : BYTE;
    Soft_Dimm : BOOL;
    Rst_Out : BOOL;
    OUT_LinearScaleMin : INT;
    OUT_LinearScaleMax : INT;
  END_VAR
                  THIS^.T_Debounce:=T_Debounce;
THIS^.T_Reconfig:=T_Reconfig;
THIS^.T_On_Max:=T_On_Max;
THIS^.T_Dimm_Start:=T_Dimm_Start;
THIS^.T_Dimm:=T_Dimm;
THIS^.Min_On:=Min_On;
THIS^.Max_On:=Max_On;
THIS^.Soft_Dimm:=Soft_Dimm;
THIS^.Rst_Out:=Rst_Out;
THIS^.OUT_LinearScaleMin:=OUT_LinearScaleMin;
THIS^.OUT_LinearScaleMax:=OUT_LinearScaleMax;
                
END_METHOD

METHOD PublishReceived : BOOL
  VAR_INPUT
    Data : MQTT.CALLBACK_DATA;  (* Collection of recived Data *)
  END_VAR
                  //first check if Mqtt is initialized, otherwise do nothing
IF NOT(InitMqttDone) THEN
	//mark the interface call from the collector as done
	PublishReceived := TRUE;
//check if the packet is for this FB
ELSIF CommonTypesAndFunctions.StrEquals(str1:= ADR(MQTTSubscribeTopic), str2:= Data.TopicOut) THEN
	//mark the interface call from the collector as done
	PublishReceived := TRUE;
	//now process the data
	IF CommonTypesAndFunctions.StrEquals(str1:= Data.PayloadString, str2:= ADR('TRUE')) THEN
		MqttHighRequest := TRUE;
	ELSIF CommonTypesAndFunctions.StrEquals(str1:= Data.PayloadString, str2:= ADR('FALSE')) THEN
		MqttLowRequest := TRUE;
	ELSIF OSCAT_BASIC.IS_CC(str:= Data.PayloadString^,cmp:='0123456789.') AND THIS^.PRIO_HIGH = FALSE THEN
		THIS^.OUT_Internal:=STRING_TO_BYTE(Data.PayloadString^);
	END_IF
END_IF 
                
END_METHOD
END_FUNCTION_BLOCK

{attribute 'reflection'}
FUNCTION_BLOCK FB_OUTPUT_SWITCH_MQTT IMPLEMENTS MQTT.MQTT_SUBSCRIBE_CALLBACK
  VAR_INPUT
    PRIO_HIGH : BOOL := FALSE;
    PRIO_LOW : BOOL := FALSE;
    TOGGLE : BOOL := FALSE;
  END_VAR
  VAR_OUTPUT
    OUT : BOOL;
  END_VAR
  VAR
    {attribute 'instance-path'}
    {attribute 'noinit'}
    InstanceName : STRING;  (* object's full instance name *)
    Startup : BOOL := TRUE;
    InitMqttDone : BOOL;
    MqttPublishTopicPrefix : POINTER TO STRING;
    MqttPublishTopicSuffix : STRING(50);
    MQTTSubscribeTopic : STRING(50);
    pMqttPublishQueue : POINTER TO FB_MqttPublishQueue;
    MqttHighRequest : BOOL;
    MqttLowRequest : BOOL;
  END_VAR
  VAR PERSISTENT
    PreviousState : BOOL;  (* To retain output state through powercycles *)
  END_VAR

            IF Startup THEN
	OUT := PreviousState;
END_IF

IF PRIO_HIGH THEN
	OUT:=TRUE;
ELSIF(PRIO_LOW AND NOT (PRIO_HIGH)) THEN
	OUT:= FALSE;
ELSIF MqttHighRequest THEN
	OUT:= TRUE;
	MqttHighRequest := FALSE;
	MqttLowRequest := FALSE;
ELSIF MqttLowRequest THEN
	OUT:= FALSE;
	MqttHighRequest := FALSE;
	MqttLowRequest := FALSE;
ELSIF(TOGGLE) THEN
	OUT:=NOT(OUT);
END_IF;

IF ((PreviousState <> OUT) OR Startup) AND InitMqttDone THEN
	pMqttPublishQueue^.AddMessage(
		Payload := BOOL_TO_STRING(OUT),
		Topic := CONCAT(MqttPublishTopicPrefix^, MqttPublishTopicSuffix),
		Qos := MQTT.QoS.ExactlyOnce,
		MqttRetain := TRUE
	);	
	Startup:=FALSE;
END_IF	

PreviousState := OUT;
          

METHOD InitMqtt
  VAR_INPUT
    MQTTPublishPrefix : POINTER TO STRING;
    MQTTSubscribePrefix : POINTER TO STRING;
    pMqttPublishQueue : POINTER TO FB_MqttPublishQueue;
    pMqttCallbackCollector : POINTER TO MQTT.CallbackCollector;
  END_VAR
  VAR
    InstanceNamePt : POINTER TO STRING;
  END_VAR
                  THIS^.pMqttPublishQueue := pMqttPublishQueue;
THIS^.MqttPublishTopicPrefix := MQTTPublishPrefix;

InstanceNamePt := CommonTypesAndFunctions.FindLastDot(ADR(THIS^.InstanceName)) + 1;
THIS^.MqttPublishTopicSuffix := InstanceNamePt^;
THIS^.MQTTSubscribeTopic := CONCAT(MQTTSubscribePrefix^ ,THIS^.MqttPublishTopicSuffix);

// register the FB agains the collector so mqtt events can be received
pMqttCallbackCollector^.put(instance:= THIS^);

InitMqttDone := TRUE;
                
END_METHOD

METHOD PublishReceived : BOOL
  VAR_INPUT
    Data : MQTT.CALLBACK_DATA;  (* Collection of recived Data *)
  END_VAR
                  //first check if Mqtt is initialized, otherwise do nothing
IF NOT(InitMqttDone) THEN
	//mark the interface call from the collector as done
	PublishReceived := TRUE;
//check if the packet is for this FB
ELSIF CommonTypesAndFunctions.StrEquals(str1:= ADR(MQTTSubscribeTopic), str2:= Data.TopicOut) THEN
	//mark the interface call from the collector as done
	PublishReceived := TRUE;
	//now process the data
	IF CommonTypesAndFunctions.StrEquals(str1:= Data.PayloadString, str2:= ADR('TRUE')) THEN
		MqttHighRequest := TRUE;
	END_IF
	IF CommonTypesAndFunctions.StrEquals(str1:= Data.PayloadString, str2:= ADR('FALSE')) THEN
		MqttLowRequest := TRUE;
	END_IF
END_IF 
                
END_METHOD
END_FUNCTION_BLOCK

FUNCTION_BLOCK FB_RS485_BUSCONTROLLER
  VAR_OUTPUT
    BusOcupied : BOOL := TRUE;  (* Set this to True by default at startup to allow for some RS485 devices to boot up at power interuptions *)
  END_VAR
  VAR
    StartupDelay : TIME := TIME#5s0ms;  (* Amount of time that should be waited on PLC startup to start using the RS485 bus *)
    SilenceTime : TIME := TIME#20ms;  (* This is the silence time between two requests *)
    Startup : BOOL := TRUE;  (* Used to detect startup *)
    tonDelay : TON;  (* To manage silence time and startup delay *)
    devices : ARRAY[0..31] OF RS485Device;  (* collection of devices on the bus *)
    devicesCount : INT := 0;  (* total number of devices registred on the bus *)
    selectedDevice : INT := 0;  (* index of the active device on the bus *)
    deviceActive : BOOL;
    loopCounter : INT;
    ActiveRtuQuery : RS485_RtuQuery;
    BusTrigger : POINTER TO BOOL;
    QueryReady : Standard.F_TRIG;
    BusData : POINTER TO ARRAY[0..124] OF WORD;
    BusError : POINTER TO BOOL;
    exc : __SYSTEM.ExceptionCode;
  END_VAR

            IF Startup THEN
	tonDelay.PT := StartupDelay;
	tonDelay.IN := TRUE;
	Startup := FALSE;
END_IF

QueryReady(CLK := BusTrigger^);
BusOcupied := NOT(tonDelay.Q);
tonDelay();

// check if there's a device that requires bus time and if so, launch the query
IF busOcupied = FALSE AND devicesCount <> 0 THEN
	FOR loopCounter := 0 TO devicesCount - 1 DO
		IF devices[loopCounter].RequestBusTime() AND deviceActive = FALSE THEN
			selectedDevice := loopCounter;
			THIS^.SetBusOccupied();
			ActiveRtuQuery := devices[selectedDevice].GetRtuQuery();
			BusTrigger^ := TRUE;
		END_IF
	END_FOR;
END_IF

//watch the trigger, when completed call the FB with the data, release the bus
IF QueryReady.Q THEN
	devices[selectedDevice].ProcessDataArray(BusError, BusData);
	THIS^.ReleaseBus();
END_IF


//let the busdevices to their work
//FOR loopCounter := 0 TO devicesCount - 1 DO
//	devices[loopCounter]();
// END_FOR;
          

METHOD RegisterDevice
  VAR_INPUT
    device : RS485Device;
  END_VAR
                  IF devicesCount <> 32 THEN
	devices[devicesCount] := device;
	devicesCount := devicesCount + 1;
END_IF
                
END_METHOD

METHOD Init
  VAR_INPUT
    StartupDelay : TIME;  (* Amount of time that should be waited on PLC startup to start using the RS485 bus, can prevent errors due to devices not booted up yet *)
    SilenceTime : TIME;  (* This is the silence time between two requests *)
    BusTrigger : POINTER TO BOOL;  (* pointer to the bool that controls triggering busrequests *)
    BusData : POINTER TO ARRAY[0..124] OF WORD;
    BusError : POINTER TO BOOL;
  END_VAR
                  THIS^.StartupDelay := StartupDelay;
THIS^.SilenceTime := SilenceTime;
THIS^.BusTrigger := BusTrigger;
THIS^.BusData := BusData;
THIS^.BusError := BusError;
                
END_METHOD

METHOD SetBusOccupied
                  THIS^.tonDelay.IN := FALSE;
THIS^.deviceActive := TRUE;
                
END_METHOD

METHOD ReleaseBus
                  // Start a timer to release the bus
THIS^.tonDelay.PT := THIS^.SilenceTime;
THIS^.tonDelay.IN := TRUE;
THIS^.deviceActive := FALSE;
                
END_METHOD
END_FUNCTION_BLOCK

{attribute 'reflection'}
FUNCTION_BLOCK FB_RS485_EASTRON_SDM_POWER_MQTT IMPLEMENTS RS485Device
  VAR_OUTPUT
    ACTIVEPOWER : REAL := 0;
    DataAvailable : BOOL := FALSE;
    Error : BOOL := FALSE;
  END_VAR
  VAR
    {attribute 'instance-path'}
    {attribute 'noinit'}
    InstanceName : STRING;  (* object's full instance name *)
    Startup : BOOL := TRUE;
    InitMqttDone : BOOL;
    MqttPublishTopicPrefix : POINTER TO STRING;
    MqttPublishTopicSuffix : STRING(50);
    pMqttPublishQueue : POINTER TO FB_MqttPublishQueue;
    InitRS485Done : BOOL := FALSE;
    ActiveDevice : BOOL := FALSE;
    timerData : TON;
    isDataUpdated : BOOL := FALSE;
    DeviceType : RS485_EASTRON_SDM_Devices;
    SDM120AndSDM220RtuQuery : RS485_RtuQuery := (FunctionCode := 4, ReadAddress := 12, ReadQuantity := 2);
    SDM630RtuQuery : RS485_RtuQuery := (FunctionCode := 4, ReadAddress := 52, ReadQuantity := 2);
  END_VAR

            timerData();

IF isDataUpdated THEN
	isDataUpdated := FALSE;
	
	IF InitMqttDone THEN
		pMqttPublishQueue^.AddMessage(
			Payload := REAL_TO_STRING(ACTIVEPOWER),
			Topic := CONCAT(CONCAT(MqttPublishTopicPrefix^, MqttPublishTopicSuffix), '/ACTP' ),
			Qos := MQTT.QoS.ExactlyOnce,
			MqttRetain := FALSE
		);
	END_IF
END_IF

          

METHOD ProcessDataArray
  VAR_INPUT
    Error : POINTER TO BOOL;
    Data : POINTER TO ARRAY[0..124] OF WORD;
  END_VAR
                  THIS^.Error := Error^;
THIS^.timerData.IN := TRUE;

IF Error^ THEN
	PubMqttMessage(Suffix := '/availability', Data := 'offline');
ELSE
	PubMqttMessage(Suffix := '/availability', Data := 'online');
END_IF

IF NOT Error^ THEN
	THIS^.ACTIVEPOWER := SwapWordsToReal(Data^[0], Data^[1]);
	THIS^.isDataUpdated := TRUE;
END_IF

ActiveDevice := FALSE;




                
END_METHOD

METHOD InitRS485
  VAR_INPUT
    DataPollingInterval : TIME;
    DeviceAddress : BYTE;
    DeviceType : RS485_EASTRON_SDM_Devices;
  END_VAR
                  THIS^.timerData.PT := DataPollingInterval;
THIS^.SDM120AndSDM220RtuQuery.DeviceId := DeviceAddress;
THIS^.SDM630RtuQuery.DeviceId := DeviceAddress;
THIS^.timerData.IN := TRUE;
THIS^.DeviceType := DeviceType;

THIS^.InitRS485Done := TRUE;
                
END_METHOD

METHOD InitMqtt
  VAR_INPUT
    MQTTPublishPrefix : POINTER TO STRING;
    pMqttPublishQueue : POINTER TO FB_MqttPublishQueue;
  END_VAR
  VAR
    InstanceNamePt : POINTER TO STRING;
  END_VAR
                  THIS^.pMqttPublishQueue := pMqttPublishQueue;
THIS^.MqttPublishTopicPrefix := MQTTPublishPrefix;

InstanceNamePt := CommonTypesAndFunctions.FindLastDot(ADR(THIS^.InstanceName)) + 1;
THIS^.MqttPublishTopicSuffix := InstanceNamePt^;

THIS^.InitMqttDone := TRUE;
                
END_METHOD

METHOD RequestBusTime : BOOL
                  IF NOT InitRS485Done THEN	
	RequestBusTime := FALSE;	
ELSIF timerData.Q THEN
	RequestBusTime := TRUE;
ELSE
	RequestBusTime := FALSE;	
END_IF
                
END_METHOD

METHOD GetRtuQuery : RS485_RtuQuery
                  IF timerData.Q THEN
	THIS^.timerData.IN := FALSE;
	IF DeviceType = RS485_EASTRON_SDM_Devices.SDM120 OR  DeviceType = RS485_EASTRON_SDM_Devices.SDM220 THEN
		GetRtuQuery := THIS^.SDM120AndSDM220RtuQuery;		
	END_IF
	IF DeviceType = RS485_EASTRON_SDM_Devices.SDM630 THEN
		GetRtuQuery := THIS^.SDM630RtuQuery;		
	END_IF
END_IF
                
END_METHOD

METHOD PubMqttMessage
  VAR_INPUT
    Suffix : STRING(100);
    Data : STRING(100);
  END_VAR
                  IF InitMqttDone THEN
		pMqttPublishQueue^.AddMessage(
			Payload := Data,
			Topic := CONCAT(CONCAT(MqttPublishTopicPrefix^, MqttPublishTopicSuffix), Suffix ),
			Qos := MQTT.QoS.ExactlyOnce,
			MqttRetain := FALSE
		);
END_IF
                
END_METHOD
END_FUNCTION_BLOCK

{attribute 'reflection'}
FUNCTION_BLOCK FB_RS485_EASTRON_SDM220_MQTT IMPLEMENTS RS485Device
  VAR_OUTPUT
    VOLTAGE : REAL := 0;
    CURRENT : REAL := 0;
    ACTIVEPOWER : REAL := 0;
    APPARENT_POWER : REAL := 0;
    REACTIVE_POWER : REAL := 0;
    POWER_FACTOR : REAL := 0;
    PHASE_ANGLE : REAL := 0;
    DataAvailable1 : BOOL := FALSE;
    Error1 : BOOL := FALSE;
    FREQUENCY : REAL := 0;
    IMPORT_ACTIVE_ENERGY : REAL := 0;
    EXPORT_ACTIVE_ENERGY : REAL := 0;
    IMPORT_REACTIVE_ENERGY : REAL := 0;
    EXPORT_REACTIVE_ENERGY : REAL := 0;
    DataAvailable2 : BOOL := FALSE;
    Error2 : BOOL := FALSE;
    TOTAL_ACTIVE_ENERGY : REAL := 0;
    TOTAL_REACTIVE_ENERGY : REAL := 0;
    DataAvailable3 : BOOL := FALSE;
    Error3 : BOOL := FALSE;
  END_VAR
  VAR
    {attribute 'instance-path'}
    {attribute 'noinit'}
    InstanceName : STRING;  (* object's full instance name *)
    Startup : BOOL := TRUE;
    InitMqttDone : BOOL;
    MqttPublishTopicPrefix : POINTER TO STRING;
    MqttPublishTopicSuffix : STRING(50);
    pMqttPublishQueue : POINTER TO FB_MqttPublishQueue;
    InitRS485Done : BOOL := FALSE;
    ActiveDevice : BOOL := FALSE;
    ActiveRtuQuery : INT := 0;
    Data1RtuQuery : RS485_RtuQuery := (FunctionCode := 4, ReadAddress := 0, ReadQuantity := 40);
    Update1 : BOOL := FALSE;
    timerData1 : TON;
    Data2RtuQuery : RS485_RtuQuery := (FunctionCode := 4, ReadAddress := 70, ReadQuantity := 10);
    Update2 : BOOL := FALSE;
    timerData2 : TON;
    Data3RtuQuery : RS485_RtuQuery := (FunctionCode := 4, ReadAddress := 342, ReadQuantity := 4);
    Update3 : BOOL := FALSE;
    timerData3 : TON;
  END_VAR

            timerData1();
timerData2();
timerData3();

IF Update1 THEN
	Update1 := FALSE;
	DataAvailable1 := TRUE;
	
	IF InitMqttDone THEN
		pMqttPublishQueue^.AddMessage(
			Payload := REAL_TO_STRING(VOLTAGE),
			Topic := CONCAT(CONCAT(MqttPublishTopicPrefix^, MqttPublishTopicSuffix), '/VOLT' ),
			Qos := MQTT.QoS.ExactlyOnce,
			MqttRetain := FALSE
		);
		pMqttPublishQueue^.AddMessage(
			Payload := REAL_TO_STRING(CURRENT),
			Topic := CONCAT(CONCAT(MqttPublishTopicPrefix^, MqttPublishTopicSuffix), '/CURR' ),
			Qos := MQTT.QoS.ExactlyOnce,
			MqttRetain := FALSE
		);	
		pMqttPublishQueue^.AddMessage(
			Payload := REAL_TO_STRING(ACTIVEPOWER),
			Topic := CONCAT(CONCAT(MqttPublishTopicPrefix^, MqttPublishTopicSuffix), '/ACTP' ),
			Qos := MQTT.QoS.ExactlyOnce,
			MqttRetain := FALSE
		);
		pMqttPublishQueue^.AddMessage(
			Payload := REAL_TO_STRING(APPARENT_POWER),
			Topic := CONCAT(CONCAT(MqttPublishTopicPrefix^, MqttPublishTopicSuffix), '/APPP' ),
			Qos := MQTT.QoS.ExactlyOnce,
			MqttRetain := FALSE
		);
		pMqttPublishQueue^.AddMessage(
			Payload := REAL_TO_STRING(REACTIVE_POWER),
			Topic := CONCAT(CONCAT(MqttPublishTopicPrefix^, MqttPublishTopicSuffix), '/REAP' ),
			Qos := MQTT.QoS.ExactlyOnce,
			MqttRetain := FALSE
		);
		pMqttPublishQueue^.AddMessage(
			Payload := REAL_TO_STRING(POWER_FACTOR),
			Topic := CONCAT(CONCAT(MqttPublishTopicPrefix^, MqttPublishTopicSuffix), '/POWF' ),
			Qos := MQTT.QoS.ExactlyOnce,
			MqttRetain := FALSE
		);
		pMqttPublishQueue^.AddMessage(
			Payload := REAL_TO_STRING(PHASE_ANGLE),
			Topic := CONCAT(CONCAT(MqttPublishTopicPrefix^, MqttPublishTopicSuffix), '/PHAA' ),
			Qos := MQTT.QoS.ExactlyOnce,
			MqttRetain := FALSE
		);
	END_IF
END_IF

IF Update2 THEN
	Update2 := FALSE;
	DataAvailable2 := TRUE;
	
	IF InitMqttDone THEN
		pMqttPublishQueue^.AddMessage(
			Payload := REAL_TO_STRING(FREQUENCY),
			Topic := CONCAT(CONCAT(MqttPublishTopicPrefix^, MqttPublishTopicSuffix), '/FREQ' ),
			Qos := MQTT.QoS.ExactlyOnce,
			MqttRetain := FALSE
		);
		pMqttPublishQueue^.AddMessage(
			Payload := REAL_TO_STRING(IMPORT_ACTIVE_ENERGY),
			Topic := CONCAT(CONCAT(MqttPublishTopicPrefix^, MqttPublishTopicSuffix), '/IMAE' ),
			Qos := MQTT.QoS.ExactlyOnce,
			MqttRetain := FALSE
		);
		pMqttPublishQueue^.AddMessage(
			Payload := REAL_TO_STRING(EXPORT_ACTIVE_ENERGY),
			Topic := CONCAT(CONCAT(MqttPublishTopicPrefix^, MqttPublishTopicSuffix), '/EXAE' ),
			Qos := MQTT.QoS.ExactlyOnce,
			MqttRetain := FALSE
		);
		pMqttPublishQueue^.AddMessage(
			Payload := REAL_TO_STRING(IMPORT_REACTIVE_ENERGY),
			Topic := CONCAT(CONCAT(MqttPublishTopicPrefix^, MqttPublishTopicSuffix), '/IMRE' ),
			Qos := MQTT.QoS.ExactlyOnce,
			MqttRetain := FALSE
		);
		pMqttPublishQueue^.AddMessage(
			Payload := REAL_TO_STRING(EXPORT_REACTIVE_ENERGY),
			Topic := CONCAT(CONCAT(MqttPublishTopicPrefix^, MqttPublishTopicSuffix), '/EXRE' ),
			Qos := MQTT.QoS.ExactlyOnce,
			MqttRetain := FALSE
		);
	END_IF
END_IF

IF Update3 THEN
	Update3 := FALSE;	
	DataAvailable3 := TRUE;
	
	IF InitMqttDone THEN
		pMqttPublishQueue^.AddMessage(
			Payload := REAL_TO_STRING(TOTAL_ACTIVE_ENERGY),
			Topic := CONCAT(CONCAT(MqttPublishTopicPrefix^, MqttPublishTopicSuffix), '/TOTAE' ),
			Qos := MQTT.QoS.ExactlyOnce,
			MqttRetain := FALSE
		);
		pMqttPublishQueue^.AddMessage(
			Payload := REAL_TO_STRING(TOTAL_REACTIVE_ENERGY),
			Topic := CONCAT(CONCAT(MqttPublishTopicPrefix^, MqttPublishTopicSuffix), '/TOTRE' ),
			Qos := MQTT.QoS.ExactlyOnce,
			MqttRetain := FALSE
		);
	END_IF
END_IF
          

METHOD ProcessDataArray
  VAR_INPUT
    Error : POINTER TO BOOL;
    Data : POINTER TO ARRAY[0..124] OF WORD;
  END_VAR
                  IF Error^ THEN
	PubMqttMessage(Suffix := '/availability', Data := 'offline');
ELSE
	PubMqttMessage(Suffix := '/availability', Data := 'online');
END_IF

IF ActiveRtuQuery = 1 THEN
	THIS^.Error1 := Error^;
	THIS^.timerData1.IN := TRUE;
	IF NOT Error^ THEN
		THIS^.VOLTAGE := SwapWordsToReal(Data^[0], Data^[1]);
		THIS^.CURRENT := SwapWordsToReal(Data^[6], Data^[7]);
		THIS^.ACTIVEPOWER := SwapWordsToReal(Data^[12], Data^[13]);
		THIS^.APPARENT_POWER := SwapWordsToReal(Data^[18], Data^[19]);
		THIS^.REACTIVE_POWER := SwapWordsToReal(Data^[24], Data^[25]);
		THIS^.POWER_FACTOR := SwapWordsToReal(Data^[30], Data^[31]);
		THIS^.PHASE_ANGLE := SwapWordsToReal(Data^[36], Data^[37]);
		THIS^.Update1 := TRUE;
	END_IF
ELSIF ActiveRtuQuery = 2 THEN
	THIS^.Error2:= Error^;
	THIS^.timerData2.IN := TRUE;
	IF NOT Error^ THEN		
		THIS^.FREQUENCY := SwapWordsToReal(Data^[0], Data^[1]);
		THIS^.IMPORT_ACTIVE_ENERGY := SwapWordsToReal(Data^[2], Data^[3]);
		THIS^.EXPORT_ACTIVE_ENERGY := SwapWordsToReal(Data^[4], Data^[5]);
		THIS^.IMPORT_REACTIVE_ENERGY := SwapWordsToReal(Data^[6], Data^[7]);
		THIS^.EXPORT_REACTIVE_ENERGY := SwapWordsToReal(Data^[8], Data^[9]);
		THIS^.Update2 := TRUE;
	END_IF
ELSIF ActiveRtuQuery = 3 THEN
	THIS^.Error3 := Error^;
	THIS^.timerData3.IN := TRUE;
	IF NOT Error^ THEN
		THIS^.TOTAL_ACTIVE_ENERGY := SwapWordsToReal(Data^[0], Data^[1]);
		THIS^.TOTAL_REACTIVE_ENERGY := SwapWordsToReal(Data^[2], Data^[3]);
		THIS^.Update3 := TRUE;
	END_IF	
END_IF

ActiveRtuQuery := 0;
ActiveDevice := FALSE;




                
END_METHOD

METHOD InitRS485
  VAR_INPUT
    Data1PollingInterval : TIME;
    Data2PollingInterval : TIME;
    Data3PollingInterval : TIME;
    DeviceAddress : BYTE;
  END_VAR
                  THIS^.timerData1.PT := Data1PollingInterval;
THIS^.timerData2.PT := Data2PollingInterval;
THIS^.timerData3.PT := Data3PollingInterval;

THIS^.Data1RtuQuery.DeviceId := DeviceAddress;
THIS^.Data2RtuQuery.DeviceId := DeviceAddress;
THIS^.Data3RtuQuery.DeviceId := DeviceAddress;

THIS^.timerData1.IN := TRUE;
THIS^.timerData2.IN := TRUE;
THIS^.timerData3.IN := TRUE;

THIS^.InitRS485Done := TRUE;
                
END_METHOD

METHOD InitMqtt
  VAR_INPUT
    MQTTPublishPrefix : POINTER TO STRING;
    pMqttPublishQueue : POINTER TO FB_MqttPublishQueue;
  END_VAR
  VAR
    InstanceNamePt : POINTER TO STRING;
  END_VAR
                  THIS^.pMqttPublishQueue := pMqttPublishQueue;
THIS^.MqttPublishTopicPrefix := MQTTPublishPrefix;

InstanceNamePt := CommonTypesAndFunctions.FindLastDot(ADR(THIS^.InstanceName)) + 1;
THIS^.MqttPublishTopicSuffix := InstanceNamePt^;

THIS^.InitMqttDone := TRUE;
                
END_METHOD

METHOD RequestBusTime : BOOL
                  IF NOT InitRS485Done THEN	
	RequestBusTime := FALSE;	
ELSIF timerData1.Q OR timerData2.Q OR timerData3.Q THEN
	RequestBusTime := TRUE;	
ELSE
	RequestBusTime := FALSE;		
END_IF
                
END_METHOD

METHOD GetRtuQuery : RS485_RtuQuery
                  IF timerData1.Q THEN
	THIS^.timerData1.IN := FALSE;
	THIS^.ActiveRtuQuery := 1;
	GetRtuQuery := THIS^.Data1RtuQuery;
ELSIF timerData2.Q THEN
	THIS^.timerData2.IN := FALSE;
	THIS^.ActiveRtuQuery := 2;
	GetRtuQuery := THIS^.Data2RtuQuery;
ELSIF timerData3.Q THEN
	THIS^.timerData3.IN := FALSE;
	THIS^.ActiveRtuQuery := 3;
	GetRtuQuery := THIS^.Data3RtuQuery;	
END_IF
                
END_METHOD

METHOD PubMqttMessage
  VAR_INPUT
    Suffix : STRING(100);
    Data : STRING(100);
  END_VAR
                  IF InitMqttDone THEN
		pMqttPublishQueue^.AddMessage(
			Payload := Data,
			Topic := CONCAT(CONCAT(MqttPublishTopicPrefix^, MqttPublishTopicSuffix), Suffix ),
			Qos := MQTT.QoS.ExactlyOnce,
			MqttRetain := FALSE
		);
END_IF
                
END_METHOD
END_FUNCTION_BLOCK

{attribute 'reflection'}
FUNCTION_BLOCK FB_RS485_ESERA_1WIRE_GATEWAY_MQTT IMPLEMENTS RS485Device
  VAR
    {attribute 'instance-path'}
    {attribute 'noinit'}
    InstanceName : STRING;  (* object's full instance name *)
    InitRS485Done : BOOL := FALSE;
    DeviceAddress : BYTE;
    OwdDevices : ARRAY[1..30] OF FB_RS485_ESERA_OWD_MQTT;
    ActiveDevice : BOOL := FALSE;
    ActiveOwd : UINT := 0;
    loopCounter : UINT;
    timerData : TON;
  END_VAR

            timerData();

FOR loopCounter := 1 TO 30 DO
	OwdDevices[loopCounter]();
END_FOR
          

METHOD GetRtuQuery : RS485_RtuQuery
                  IF timerData.Q THEN
	THIS^.timerData.IN := FALSE;
	GetRtuQuery := THIS^.OwdDevices[ActiveOwd].GetRtuQuery();	
END_IF
                
END_METHOD

METHOD ProcessDataArray
  VAR_INPUT
    Error : POINTER TO BOOL;
    Data : POINTER TO ARRAY[0..124] OF WORD;
  END_VAR
                  THIS^.OwdDevices[ActiveOwd].ProcessDataArray(
	Data := Data,
	Error := Error
);
THIS^.ActiveOwd := 0;
THIS^.timerData.IN := TRUE;
                
END_METHOD

METHOD RequestBusTime : BOOL
                  IF NOT InitRS485Done OR NOT timerData.Q THEN	
	RequestBusTime := FALSE;
ELSE
	FOR loopCounter := 1 TO 30 DO
		IF OwdDevices[loopCounter].RequestBusTime() AND RequestBusTime = FALSE THEN
			THIS^.ActiveOwd := loopCounter;
			RequestBusTime := TRUE;			
		END_IF
	END_FOR
END_IF
                
END_METHOD

METHOD InitRS485
  VAR_INPUT
    DeviceAddress : BYTE;
  END_VAR
                  THIS^.DeviceAddress := DeviceAddress;
THIS^.timerData.PT := T#250MS;
THIS^.timerData.IN := TRUE;
THIS^.InitRS485Done := TRUE;
                
END_METHOD

METHOD InitMqtt
  VAR_INPUT
    MQTTPublishPrefix : POINTER TO STRING;
    pMqttPublishQueue : POINTER TO FB_MqttPublishQueue;
  END_VAR
  VAR
    InstanceNamePt : POINTER TO STRING;
  END_VAR
                  InstanceNamePt := CommonTypesAndFunctions.FindLastDot(ADR(THIS^.InstanceName)) + 1;

FOR loopCounter := 1 TO 30 DO
		OwdDevices[loopCounter].InitMqtt(
			MQTTPublishPrefix := MQTTPublishPrefix,
			MqttPublishTopicSuffix := InstanceNamePt^,
			pMqttPublishQueue := pMqttPublishQueue
		);
END_FOR
                
END_METHOD

METHOD EnableOwd : BOOL
  VAR_INPUT
    OwdNumber : UINT;
    DataPollingInterval : TIME;
  END_VAR
                  THIS^.OwdDevices[OwdNumber].InitOwd(
	DeviceAddress := THIS^.DeviceAddress,
	OwdNumber := OwdNumber,
	DataPollingInterval := DataPollingInterval
);
                
END_METHOD
END_FUNCTION_BLOCK

FUNCTION_BLOCK FB_RS485_ESERA_OWD_MQTT
  VAR_OUTPUT
    OWD_VOLTAGE : REAL := 0;
    TEMPERATURE : REAL := 0;
    HUMIDITY : REAL := 0;
    DEW_POINT : REAL := 0;
    AIR_QUALITY : REAL := 0;
    BRIGHTNESS : REAL := 0;
    DataAvailable : BOOL := FALSE;
    Error : BOOL := FALSE;
  END_VAR
  VAR
    OwdNumber : UINT;
    InitMqttDone : BOOL;
    MqttPublishTopicPrefix : POINTER TO STRING;
    MqttPublishTopicSuffix : STRING(50);
    pMqttPublishQueue : POINTER TO FB_MqttPublishQueue;
    InitOwdDone : BOOL := FALSE;
    timerData : TON;
    RtuQuery : RS485_RtuQuery := (FunctionCode := 3, ReadAddress := 100, ReadQuantity := 17);
  END_VAR

            timerData();


          

METHOD GetRtuQuery : RS485_RtuQuery
                  IF timerData.Q THEN
	THIS^.timerData.IN := FALSE;
	GetRtuQuery := THIS^.RtuQuery;	
END_IF
                
END_METHOD

METHOD ProcessDataArray
  VAR_INPUT
    Error : POINTER TO BOOL;
    Data : POINTER TO ARRAY[0..124] OF WORD;
  END_VAR
                  THIS^.timerData.IN := TRUE;

IF WORD_TO_INT(Data^[12]) <> 0 OR Error^ THEN
	THIS^.Error := TRUE;
	PubMqttMessage(Suffix := '/availability', Data := 'offline');
ELSE 	
	THIS^.Error := FALSE;
	THIS^.DataAvailable := TRUE;
	PubMqttMessage(Suffix := '/availability', Data := 'online');
END_IF

// Data handling
IF NOT Error^ AND WORD_TO_INT(Data^[12]) = 0 THEN
	IF Data^[16] = 11151 OR Data^[16] = 11152 THEN // Temperature, humidity & air quality
		ProcessTemperature(Data^[0]);		
		ProcessOwdVoltage(Data^[2]);
		ProcessHumidity(Data^[4]);
		ProcessDewPoint(Data^[6]);
		ProcessAirQuality(Data^[8]);
	ELSIF Data^[16] = 11102 OR Data^[16] = 11113 OR Data^[16] = 11120 OR Data^[16] = 11148 OR Data^[16] = 11150 OR Data^[16] = 11160 THEN // Temperature, humidity
		ProcessTemperature(Data^[0]);		
		ProcessOwdVoltage(Data^[2]);
		ProcessHumidity(Data^[4]);
		ProcessDewPoint(Data^[6]);
	ELSIF Data^[16] = 11121 OR Data^[16] = 11132 OR Data^[16] = 11134 OR Data^[16] = 11135 THEN // Temperature, humidity, brightness
		ProcessTemperature(Data^[0]);		
		ProcessOwdVoltage(Data^[2]);
		ProcessHumidity(Data^[4]);
		ProcessDewPoint(Data^[6]);
		ProcessBrigthness(Data^[8]);
	ELSIF Data^[16] = 1820  THEN // Temperature DS18B20
        ProcessTemperature(Data^[0]);
	END_IF		
END_IF
                
END_METHOD

METHOD RequestBusTime : BOOL
                  IF NOT InitOwdDone THEN	
	RequestBusTime := FALSE;	
ELSIF timerData.Q THEN
	RequestBusTime := TRUE;
ELSE
	RequestBusTime := FALSE;	
END_IF
                
END_METHOD

METHOD InitOwd
  VAR_INPUT
    DeviceAddress : BYTE;
    OwdNumber : UINT;
    DataPollingInterval : TIME;
  END_VAR
                  THIS^.RtuQuery.DeviceId := DeviceAddress;
THIS^.RtuQuery.ReadAddress := OwdNumber * 100;
THIS^.timerData.PT := DataPollingInterval;
THIS^.OwdNumber := OwdNumber;

THIS^.timerData.IN := TRUE;

THIS^.InitOwdDone := TRUE;
                
END_METHOD

METHOD InitMqtt
  VAR_INPUT
    MQTTPublishPrefix : POINTER TO STRING;
    MqttPublishTopicSuffix : STRING(255);
    pMqttPublishQueue : POINTER TO FB_MqttPublishQueue;
  END_VAR
                  THIS^.MqttPublishTopicPrefix := MQTTPublishPrefix;
THIS^.MqttPublishTopicSuffix := MqttPublishTopicSuffix;
THIS^.pMqttPublishQueue := pMqttPublishQueue;

THIS^.InitMqttDone := TRUE;
                
END_METHOD

METHOD PubMqttMessage
  VAR_INPUT
    Suffix : STRING(100);
    Data : STRING(100);
  END_VAR
                  IF InitMqttDone THEN
		pMqttPublishQueue^.AddMessage(
			Payload := Data,
			Topic := CONCAT(CONCAT(CONCAT(CONCAT(MqttPublishTopicPrefix^, MqttPublishTopicSuffix), '/OWD/'), UINT_TO_STRING(OwdNumber)), Suffix ),
			Qos := MQTT.QoS.ExactlyOnce,
			MqttRetain := FALSE
		);
END_IF
                
END_METHOD

METHOD ProcessTemperature
  VAR_INPUT
    Data : WORD;
  END_VAR
                  THIS^.TEMPERATURE := WORD_TO_REAL(Data) / 100;
PubMqttMessage(Suffix := '/TEMP', Data := REAL_TO_STRING(TEMPERATURE));
                
END_METHOD

METHOD ProcessOwdVoltage
  VAR_INPUT
    Data : WORD;
  END_VAR
                  THIS^.OWD_VOLTAGE := WORD_TO_REAL(Data) / 100;
PubMqttMessage(Suffix := '/OWDV', Data := REAL_TO_STRING(OWD_VOLTAGE));
                
END_METHOD

METHOD ProcessHumidity
  VAR_INPUT
    Data : WORD;
  END_VAR
                  THIS^.HUMIDITY := WORD_TO_REAL(Data) / 100;
PubMqttMessage(Suffix := '/HUM', Data := REAL_TO_STRING(HUMIDITY));
                
END_METHOD

METHOD ProcessDewPoint
  VAR_INPUT
    Data : WORD;
  END_VAR
                  THIS^.DEW_POINT := WORD_TO_REAL(Data) / 100;
PubMqttMessage(Suffix := '/DEWP', Data := REAL_TO_STRING(DEW_POINT));
                
END_METHOD

METHOD ProcessAirQuality
  VAR_INPUT
    Data : WORD;
  END_VAR
                  THIS^.AIR_QUALITY := WORD_TO_REAL(Data) / 100;
PubMqttMessage(Suffix := '/AIRQ', Data := REAL_TO_STRING(AIR_QUALITY));
                
END_METHOD

METHOD ProcessBrigthness
  VAR_INPUT
    Data : WORD;
  END_VAR
                  THIS^.BRIGHTNESS := WORD_TO_REAL(Data) / 100;
PubMqttMessage(Suffix := '/BNESS', Data := REAL_TO_STRING(BRIGHTNESS));
                
END_METHOD
END_FUNCTION_BLOCK

{attribute 'reflection'}
FUNCTION_BLOCK FB_VIRTUAL_BOOL_MQTT IMPLEMENTS MQTT.MQTT_SUBSCRIBE_CALLBACK
  VAR_INPUT
    IN : BOOL;
  END_VAR
  VAR_OUTPUT
    OUT : BOOL;
  END_VAR
  VAR
    {attribute 'instance-path'}
    {attribute 'noinit'}
    InstanceName : STRING;  (* object's full instance name *)
    Startup : BOOL := TRUE;
    InitMqttDone : BOOL;
    MqttPublishTopicPrefix : POINTER TO STRING;
    MqttPublishTopicSuffix : STRING(50);
    MQTTSubscribeTopic : STRING(50);
    pMqttPublishQueue : POINTER TO FB_MqttPublishQueue;
    MqttQos : MQTT.QoS;
    MqttRetain : BOOL;
    UpdateFlag : BOOL;
    VirtualMode : VIRTUAL_MODES;
    DefaultValue : BOOL;
    SetDefaultValueStartup : BOOL;
    PublishAtStartup : BOOL;
    UsePersistentAtStartup : BOOL;
    ConfirmReceival : BOOL;
    MqttMessageReceived : BOOL;
    PreviousIn : BOOL;
  END_VAR
  VAR PERSISTENT
    PreviousState : BOOL;  (* To retain output state through powercycles *)
  END_VAR

            IF VirtualMode = VIRTUAL_MODES.Output THEN
	IF (Startup AND PublishAtStartup) OR (UpdateFlag OR IN <> PreviousIn) AND InitMqttDone THEN
	pMqttPublishQueue^.AddMessage(
		Payload := BOOL_TO_STRING(IN),
		Topic := CONCAT(MqttPublishTopicPrefix^, MqttPublishTopicSuffix),
		Qos := MqttQos,
		MqttRetain := MqttRetain
	);
	Startup:=FALSE;
	UpdateFlag := FALSE;
	PreviousIn := IN;
	END_IF
ELSIF VirtualMode = VIRTUAL_MODES.Input THEN
	IF Startup AND SetDefaultValueStartup THEN
		OUT := DefaultValue;
	ELSIF UsePersistentAtStartup THEN
		OUT := PreviousState;
	END_IF	
	
	IF ((Startup AND PublishAtStartup) OR (ConfirmReceival AND MqttMessageReceived)) AND InitMqttDone THEN
	pMqttPublishQueue^.AddMessage(
		Payload := BOOL_TO_STRING(OUT),
		Topic := CONCAT(MqttPublishTopicPrefix^, MqttPublishTopicSuffix),
		Qos := MqttQos,
		MqttRetain := MqttRetain
	);
	Startup:=FALSE;
	MqttMessageReceived := FALSE;
	PreviousState:=OUT;
	END_IF		
	
END_IF
          

METHOD InitMqtt
  VAR_INPUT
    MQTTPublishPrefix : POINTER TO STRING;
    MQTTSubscribePrefix : POINTER TO STRING;
    pMqttPublishQueue : POINTER TO FB_MqttPublishQueue;
    pMqttCallbackCollector : POINTER TO MQTT.CallbackCollector;
    MqttQos : MQTT.QoS;
    MqttRetain : BOOL;
  END_VAR
  VAR
    InstanceNamePt : POINTER TO STRING;
  END_VAR
                  THIS^.pMqttPublishQueue := pMqttPublishQueue;
THIS^.MqttPublishTopicPrefix := MQTTPublishPrefix;

InstanceNamePt := CommonTypesAndFunctions.FindLastDot(ADR(THIS^.InstanceName)) + 1;
THIS^.MqttPublishTopicSuffix := InstanceNamePt^;
THIS^.MQTTSubscribeTopic := CONCAT(MQTTSubscribePrefix^ ,THIS^.MqttPublishTopicSuffix);

// register the FB agains the collector so mqtt events can be received
pMqttCallbackCollector^.put(instance:= THIS^);

THIS^.MqttQos:=MqttQos;
THIS^.MqttRetain:=MqttRetain;

InitMqttDone := TRUE;
                
END_METHOD

METHOD PublishReceived : BOOL
  VAR_INPUT
    Data : MQTT.CALLBACK_DATA;  (* Collection of recived Data *)
  END_VAR
                  //first check if Mqtt is initialized and FB in input mode, otherwise do nothing
IF NOT(InitMqttDone) AND VirtualMode <> VIRTUAL_MODES.Input THEN
	//mark the interface call from the collector as done
	PublishReceived := TRUE;
//check if the packet is for this FB
ELSIF CommonTypesAndFunctions.StrEquals(str1:= ADR(MQTTSubscribeTopic), str2:= Data.TopicOut) THEN
	//mark the interface call from the collector as done
	PublishReceived := TRUE;
	//process the data
	IF CommonTypesAndFunctions.StrEquals(str1:= Data.PayloadString, str2:= ADR('TRUE')) THEN
		THIS^.OUT := TRUE;
		MqttMessageReceived := TRUE;
	END_IF
	IF CommonTypesAndFunctions.StrEquals(str1:= Data.PayloadString, str2:= ADR('FALSE')) THEN
		THIS^.OUT := FALSE;
		MqttMessageReceived := TRUE;
	END_IF
END_IF 
                
END_METHOD

METHOD ConfigureFunctionBlockAsVirtualInput : BOOL
  VAR_INPUT
    DefaultValue : BOOL;
    SetDefaultValueStartup : BOOL;
    PublishAtStartup : BOOL;
    UsePersistentAtStartup : BOOL;
    ConfirmReceival : BOOL;
  END_VAR
                  THIS^.DefaultValue:=DefaultValue;
THIS^.SetDefaultValueStartup:=SetDefaultValueStartup;
THIS^.PublishAtStartup:=PublishAtStartup;
THIS^.UsePersistentAtStartup:=UsePersistentAtStartup;
THIS^.ConfirmReceival:=ConfirmReceival;
THIS^.VirtualMode:=VIRTUAL_MODES.Input;
                
END_METHOD

METHOD SetValue : BOOL
  VAR_INPUT
    Value : BOOL;
  END_VAR
                  THIS^.OUT:=Value;
THIS^.UpdateFlag:=TRUE;
                
END_METHOD

METHOD ConfigureFunctionBlockAsVirtualOutput : BOOL
  VAR_INPUT
    PublishAtStartup : BOOL;
  END_VAR
                  THIS^.PublishAtStartup:=PublishAtStartup;
THIS^.VirtualMode:=VIRTUAL_MODES.Output;
                
END_METHOD
END_FUNCTION_BLOCK

{attribute 'reflection'}
FUNCTION_BLOCK FB_VIRTUAL_INT_MQTT IMPLEMENTS MQTT.MQTT_SUBSCRIBE_CALLBACK
  VAR_INPUT
    IN : INT;
  END_VAR
  VAR_OUTPUT
    OUT : INT;
  END_VAR
  VAR
    {attribute 'instance-path'}
    {attribute 'noinit'}
    InstanceName : STRING;  (* object's full instance name *)
    Startup : BOOL := TRUE;
    InitMqttDone : BOOL;
    MqttPublishTopicPrefix : POINTER TO STRING;
    MqttPublishTopicSuffix : STRING(50);
    MQTTSubscribeTopic : STRING(50);
    pMqttPublishQueue : POINTER TO FB_MqttPublishQueue;
    MqttQos : MQTT.QoS;
    MqttRetain : BOOL;
    UpdateFlag : BOOL;
    VirtualMode : VIRTUAL_MODES;
    DefaultValue : INT;
    SetDefaultValueStartup : BOOL;
    PublishAtStartup : BOOL;
    UsePersistentAtStartup : BOOL;
    ConfirmReceival : BOOL;
    MqttMessageReceived : BOOL;
    PreviousIn : INT;
  END_VAR
  VAR PERSISTENT
    PreviousState : INT;  (* To retain output state through powercycles *)
  END_VAR

            IF VirtualMode = VIRTUAL_MODES.Output THEN
	IF (Startup AND PublishAtStartup) OR (UpdateFlag OR IN <> PreviousIn) AND InitMqttDone THEN
	pMqttPublishQueue^.AddMessage(
		Payload := INT_TO_STRING(IN),
		Topic := CONCAT(MqttPublishTopicPrefix^, MqttPublishTopicSuffix),
		Qos := MqttQos,
		MqttRetain := MqttRetain
	);
	Startup:=FALSE;
	UpdateFlag := FALSE;
	PreviousIn := IN;
	END_IF
ELSIF VirtualMode = VIRTUAL_MODES.Input THEN
	IF Startup AND SetDefaultValueStartup THEN
		OUT := DefaultValue;
	ELSIF UsePersistentAtStartup THEN
		OUT := PreviousState;
	END_IF	
	
	IF ((Startup AND PublishAtStartup) OR (ConfirmReceival AND MqttMessageReceived)) AND InitMqttDone THEN
	pMqttPublishQueue^.AddMessage(
		Payload := INT_TO_STRING(OUT),
		Topic := CONCAT(MqttPublishTopicPrefix^, MqttPublishTopicSuffix),
		Qos := MqttQos,
		MqttRetain := MqttRetain
	);
	Startup:=FALSE;
	MqttMessageReceived := FALSE;
	PreviousState:=OUT;
	END_IF		
	
END_IF
          

METHOD ConfigureFunctionBlockAsVirtualOutput : BOOL
  VAR_INPUT
    PublishAtStartup : BOOL;
  END_VAR
                  THIS^.PublishAtStartup:=PublishAtStartup;
THIS^.VirtualMode:=VIRTUAL_MODES.Output;
                
END_METHOD

METHOD InitMqtt
  VAR_INPUT
    MQTTPublishPrefix : POINTER TO STRING;
    MQTTSubscribePrefix : POINTER TO STRING;
    pMqttPublishQueue : POINTER TO FB_MqttPublishQueue;
    pMqttCallbackCollector : POINTER TO MQTT.CallbackCollector;
    MqttQos : MQTT.QoS;
    MqttRetain : BOOL;
  END_VAR
  VAR
    InstanceNamePt : POINTER TO STRING;
  END_VAR
                  THIS^.pMqttPublishQueue := pMqttPublishQueue;
THIS^.MqttPublishTopicPrefix := MQTTPublishPrefix;

InstanceNamePt := CommonTypesAndFunctions.FindLastDot(ADR(THIS^.InstanceName)) + 1;
THIS^.MqttPublishTopicSuffix := InstanceNamePt^;
THIS^.MQTTSubscribeTopic := CONCAT(MQTTSubscribePrefix^ ,THIS^.MqttPublishTopicSuffix);

// register the FB agains the collector so mqtt events can be received
pMqttCallbackCollector^.put(instance:= THIS^);

THIS^.MqttQos:=MqttQos;
THIS^.MqttRetain:=MqttRetain;

InitMqttDone := TRUE;
                
END_METHOD

METHOD PublishReceived : BOOL
  VAR_INPUT
    Data : MQTT.CALLBACK_DATA;  (* Collection of recived Data *)
  END_VAR
                  //first check if Mqtt is initialized and FB in input mode, otherwise do nothing
IF NOT(InitMqttDone) AND VirtualMode <> VIRTUAL_MODES.Input THEN
	//mark the interface call from the collector as done
	PublishReceived := TRUE;
//check if the packet is for this FB
ELSIF CommonTypesAndFunctions.StrEquals(str1:= ADR(MQTTSubscribeTopic), str2:= Data.TopicOut) THEN
	//mark the interface call from the collector as done
	PublishReceived := TRUE;
	//process the data
	IF OSCAT_BASIC.IS_NUM(str:= Data.PayloadString^) THEN
		THIS^.OUT := STRING_TO_INT(Data.PayloadString^);	
		MqttMessageReceived := TRUE;	
	END_IF
END_IF 
                
END_METHOD

METHOD ConfigureFunctionBlockAsVirtualInput : BOOL
  VAR_INPUT
    DefaultValue : INT;
    SetDefaultValueStartup : BOOL;
    PublishAtStartup : BOOL;
    UsePersistentAtStartup : BOOL;
    ConfirmReceival : BOOL;
  END_VAR
                  THIS^.DefaultValue:=DefaultValue;
THIS^.SetDefaultValueStartup:=SetDefaultValueStartup;
THIS^.PublishAtStartup:=PublishAtStartup;
THIS^.UsePersistentAtStartup:=UsePersistentAtStartup;
THIS^.ConfirmReceival:=ConfirmReceival;
THIS^.VirtualMode:=VIRTUAL_MODES.Input;
                
END_METHOD

METHOD SetValue : BOOL
  VAR_INPUT
    Value : INT;
  END_VAR
                  THIS^.OUT:=Value;
THIS^.UpdateFlag:=TRUE;
                
END_METHOD
END_FUNCTION_BLOCK

{attribute 'reflection'}
FUNCTION_BLOCK FB_VIRTUAL_REAL_MQTT IMPLEMENTS MQTT.MQTT_SUBSCRIBE_CALLBACK
  VAR_INPUT
    IN : REAL;
  END_VAR
  VAR_OUTPUT
    OUT : REAL;
  END_VAR
  VAR
    {attribute 'instance-path'}
    {attribute 'noinit'}
    InstanceName : STRING;  (* object's full instance name *)
    Startup : BOOL := TRUE;
    InitMqttDone : BOOL;
    MqttPublishTopicPrefix : POINTER TO STRING;
    MqttPublishTopicSuffix : STRING(50);
    MQTTSubscribeTopic : STRING(50);
    pMqttPublishQueue : POINTER TO FB_MqttPublishQueue;
    MqttQos : MQTT.QoS;
    MqttRetain : BOOL;
    UpdateFlag : BOOL;
    VirtualMode : VIRTUAL_MODES;
    DefaultValue : REAL;
    SetDefaultValueStartup : BOOL;
    PublishAtStartup : BOOL;
    UsePersistentAtStartup : BOOL;
    ConfirmReceival : BOOL;
    MqttMessageReceived : BOOL;
    PreviousIn : REAL;
  END_VAR
  VAR PERSISTENT
    PreviousState : REAL;  (* To retain output state through powercycles *)
  END_VAR

            IF VirtualMode = VIRTUAL_MODES.Output THEN
	IF (Startup AND PublishAtStartup) OR (UpdateFlag OR IN <> PreviousIn) AND InitMqttDone THEN
	pMqttPublishQueue^.AddMessage(
		Payload := REAL_TO_STRING(IN),
		Topic := CONCAT(MqttPublishTopicPrefix^, MqttPublishTopicSuffix),
		Qos := MqttQos,
		MqttRetain := MqttRetain
	);
	Startup:=FALSE;
	UpdateFlag := FALSE;
	PreviousIn := IN;
	END_IF
ELSIF VirtualMode = VIRTUAL_MODES.Input THEN
	IF Startup AND SetDefaultValueStartup THEN
		OUT := DefaultValue;
	ELSIF UsePersistentAtStartup THEN
		OUT := PreviousState;
	END_IF	
	
	IF ((Startup AND PublishAtStartup) OR (ConfirmReceival AND MqttMessageReceived)) AND InitMqttDone THEN
	pMqttPublishQueue^.AddMessage(
		Payload := REAL_TO_STRING(OUT),
		Topic := CONCAT(MqttPublishTopicPrefix^, MqttPublishTopicSuffix),
		Qos := MqttQos,
		MqttRetain := MqttRetain
	);
	Startup:=FALSE;
	MqttMessageReceived := FALSE;
	PreviousState:=OUT;
	END_IF		
	
END_IF
          

METHOD ConfigureFunctionBlockAsVirtualOutput : BOOL
  VAR_INPUT
    PublishAtStartup : BOOL;
  END_VAR
                  THIS^.PublishAtStartup:=PublishAtStartup;
THIS^.VirtualMode:=VIRTUAL_MODES.Output;
                
END_METHOD

METHOD InitMqtt
  VAR_INPUT
    MQTTPublishPrefix : POINTER TO STRING;
    MQTTSubscribePrefix : POINTER TO STRING;
    pMqttPublishQueue : POINTER TO FB_MqttPublishQueue;
    pMqttCallbackCollector : POINTER TO MQTT.CallbackCollector;
    MqttQos : MQTT.QoS;
    MqttRetain : BOOL;
  END_VAR
  VAR
    InstanceNamePt : POINTER TO STRING;
  END_VAR
                  THIS^.pMqttPublishQueue := pMqttPublishQueue;
THIS^.MqttPublishTopicPrefix := MQTTPublishPrefix;

InstanceNamePt := CommonTypesAndFunctions.FindLastDot(ADR(THIS^.InstanceName)) + 1;
THIS^.MqttPublishTopicSuffix := InstanceNamePt^;
THIS^.MQTTSubscribeTopic := CONCAT(MQTTSubscribePrefix^ ,THIS^.MqttPublishTopicSuffix);

// register the FB agains the collector so mqtt events can be received
pMqttCallbackCollector^.put(instance:= THIS^);

THIS^.MqttQos:=MqttQos;
THIS^.MqttRetain:=MqttRetain;

InitMqttDone := TRUE;
                
END_METHOD

METHOD PublishReceived : BOOL
  VAR_INPUT
    Data : MQTT.CALLBACK_DATA;  (* Collection of recived Data *)
  END_VAR
                  //first check if Mqtt is initialized and FB in input mode, otherwise do nothing
IF NOT(InitMqttDone) AND VirtualMode <> VIRTUAL_MODES.Input THEN
	//mark the interface call from the collector as done
	PublishReceived := TRUE;
//check if the packet is for this FB
ELSIF CommonTypesAndFunctions.StrEquals(str1:= ADR(MQTTSubscribeTopic), str2:= Data.TopicOut) THEN
	//mark the interface call from the collector as done
	PublishReceived := TRUE;
	//process the data
	THIS^.OUT := STRING_TO_REAL(Data.PayloadString^);	
	MqttMessageReceived := TRUE;	
END_IF 
                
END_METHOD

METHOD ConfigureFunctionBlockAsVirtualInput : BOOL
  VAR_INPUT
    DefaultValue : REAL;
    SetDefaultValueStartup : BOOL;
    PublishAtStartup : BOOL;
    UsePersistentAtStartup : BOOL;
    ConfirmReceival : BOOL;
  END_VAR
                  THIS^.DefaultValue:=DefaultValue;
THIS^.SetDefaultValueStartup:=SetDefaultValueStartup;
THIS^.PublishAtStartup:=PublishAtStartup;
THIS^.UsePersistentAtStartup:=UsePersistentAtStartup;
THIS^.ConfirmReceival:=ConfirmReceival;
THIS^.VirtualMode:=VIRTUAL_MODES.Input;
                
END_METHOD

METHOD SetValue : BOOL
  VAR_INPUT
    Value : REAL;
  END_VAR
                  THIS^.OUT:=Value;
THIS^.UpdateFlag:=TRUE;
                
END_METHOD
END_FUNCTION_BLOCK

{attribute 'reflection'}
FUNCTION_BLOCK FB_VIRTUAL_STRING_MQTT IMPLEMENTS MQTT.MQTT_SUBSCRIBE_CALLBACK
  VAR_INPUT
    IN : STRING;
  END_VAR
  VAR_OUTPUT
    OUT : STRING;
  END_VAR
  VAR
    {attribute 'instance-path'}
    {attribute 'noinit'}
    InstanceName : STRING;  (* object's full instance name *)
    Startup : BOOL := TRUE;
    InitMqttDone : BOOL;
    MqttPublishTopicPrefix : POINTER TO STRING;
    MqttPublishTopicSuffix : STRING(50);
    MQTTSubscribeTopic : STRING(50);
    pMqttPublishQueue : POINTER TO FB_MqttPublishQueue;
    MqttQos : MQTT.QoS;
    MqttRetain : BOOL;
    UpdateFlag : BOOL;
    VirtualMode : VIRTUAL_MODES;
    DefaultValue : STRING;
    SetDefaultValueStartup : BOOL;
    PublishAtStartup : BOOL;
    UsePersistentAtStartup : BOOL;
    ConfirmReceival : BOOL;
    MqttMessageReceived : BOOL;
    PreviousIn : STRING;
  END_VAR
  VAR PERSISTENT
    PreviousState : STRING;  (* To retain output state through powercycles *)
  END_VAR

            IF VirtualMode = VIRTUAL_MODES.Output THEN
	IF (Startup AND PublishAtStartup) OR (UpdateFlag OR IN <> PreviousIn) AND InitMqttDone THEN
	pMqttPublishQueue^.AddMessage(
		Payload := IN,
		Topic := CONCAT(MqttPublishTopicPrefix^, MqttPublishTopicSuffix),
		Qos := MqttQos,
		MqttRetain := MqttRetain
	);
	Startup:=FALSE;
	UpdateFlag := FALSE;
	PreviousIn := IN;
	END_IF
ELSIF VirtualMode = VIRTUAL_MODES.Input THEN
	IF Startup AND SetDefaultValueStartup THEN
		OUT := DefaultValue;
	ELSIF UsePersistentAtStartup THEN
		OUT := PreviousState;
	END_IF	
	
	IF ((Startup AND PublishAtStartup) OR (ConfirmReceival AND MqttMessageReceived)) AND InitMqttDone THEN
	pMqttPublishQueue^.AddMessage(
		Payload := OUT,
		Topic := CONCAT(MqttPublishTopicPrefix^, MqttPublishTopicSuffix),
		Qos := MqttQos,
		MqttRetain := MqttRetain
	);
	Startup:=FALSE;
	MqttMessageReceived := FALSE;
	PreviousState:=OUT;
	END_IF		
	
END_IF
          

METHOD InitMqtt
  VAR_INPUT
    MQTTPublishPrefix : POINTER TO STRING;
    MQTTSubscribePrefix : POINTER TO STRING;
    pMqttPublishQueue : POINTER TO FB_MqttPublishQueue;
    pMqttCallbackCollector : POINTER TO MQTT.CallbackCollector;
    MqttQos : MQTT.QoS;
    MqttRetain : BOOL;
  END_VAR
  VAR
    InstanceNamePt : POINTER TO STRING;
  END_VAR
                  THIS^.pMqttPublishQueue := pMqttPublishQueue;
THIS^.MqttPublishTopicPrefix := MQTTPublishPrefix;

InstanceNamePt := CommonTypesAndFunctions.FindLastDot(ADR(THIS^.InstanceName)) + 1;
THIS^.MqttPublishTopicSuffix := InstanceNamePt^;
THIS^.MQTTSubscribeTopic := CONCAT(MQTTSubscribePrefix^ ,THIS^.MqttPublishTopicSuffix);

// register the FB agains the collector so mqtt events can be received
pMqttCallbackCollector^.put(instance:= THIS^);

THIS^.MqttQos:=MqttQos;
THIS^.MqttRetain:=MqttRetain;

InitMqttDone := TRUE;
                
END_METHOD

METHOD PublishReceived : BOOL
  VAR_INPUT
    Data : MQTT.CALLBACK_DATA;  (* Collection of recived Data *)
  END_VAR
                  //first check if Mqtt is initialized and FB in input mode, otherwise do nothing
IF NOT(InitMqttDone) AND VirtualMode <> VIRTUAL_MODES.Input THEN
	//mark the interface call from the collector as done
	PublishReceived := TRUE;
//check if the packet is for this FB
ELSIF CommonTypesAndFunctions.StrEquals(str1:= ADR(MQTTSubscribeTopic), str2:= Data.TopicOut) THEN
	//mark the interface call from the collector as done
	PublishReceived := TRUE;
	//process the data
	THIS^.OUT := Data.PayloadString^;	
	MqttMessageReceived := TRUE;
END_IF 
                
END_METHOD

METHOD ConfigureFunctionBlockAsVirtualInput : BOOL
  VAR_INPUT
    DefaultValue : STRING;
    SetDefaultValueStartup : BOOL;
    PublishAtStartup : BOOL;
    UsePersistentAtStartup : BOOL;
    ConfirmReceival : BOOL;
  END_VAR
                  THIS^.DefaultValue:=DefaultValue;
THIS^.SetDefaultValueStartup:=SetDefaultValueStartup;
THIS^.PublishAtStartup:=PublishAtStartup;
THIS^.UsePersistentAtStartup:=UsePersistentAtStartup;
THIS^.ConfirmReceival:=ConfirmReceival;
THIS^.VirtualMode:=VIRTUAL_MODES.Input;
                
END_METHOD

METHOD SetValue : BOOL
  VAR_INPUT
    Value : STRING;
  END_VAR
                  THIS^.OUT:=Value;
THIS^.UpdateFlag:=TRUE;
                
END_METHOD

METHOD ConfigureFunctionBlockAsVirtualOutput : BOOL
  VAR_INPUT
    PublishAtStartup : BOOL;
  END_VAR
                  THIS^.PublishAtStartup:=PublishAtStartup;
THIS^.VirtualMode:=VIRTUAL_MODES.Output;
                
END_METHOD
END_FUNCTION_BLOCK

FUNCTION_BLOCK RMP_B
  VAR_INPUT
    SET : BOOL;
    PT : TIME;
    E : BOOL := TRUE;
    UP : BOOL := TRUE;
    RST : BOOL;
  END_VAR
  VAR_OUTPUT
    OUT : BYTE;
    BUSY : BOOL;
    HIGH : BOOL;
    LOW : BOOL;
  END_VAR
  VAR
    rmp : _RMP_B;
  END_VAR

            (* generate ramp *)
rmp(dir := UP, E := E, TR := PT, rmp := out);

(* set or reset operation *)
IF RST THEN
	out := 0;
ELSIF SET THEN
	out := 255;
END_IF;

(* checks for outputs stable and reset or set busy flag *)
low := out = 0;
high := out = 255;
busy := NOT (low OR high) AND E;


(* revision history

hm 5.10.2006	rev 1.1
	added busy output
hm 17.1.2007	rev 1.2
	renamed input ud to up for better usability
	deleted unused variable step

hm	17.9.2007		rev 1.3
	replaced time() with t_plc_ms() for compatibility reasons

hm	28. sep 2007	rev 1.4
	added outputs on and off
	busy is now disabled while en is false
	new coding for higher accuracy and performance

hm	5. oct 2007	rev 1.5
	added statements to allow for PT to be t#0s output jumps to max or min immediately

hm	25. dec 2007	rev 1.6
	improved code for better performance

hm	16. oct. 2008	rev 1.7
	improved code for better performance

hm	18. oct. 2008	rev 1.8
	added type conversion to avoid warnings
	changed input en to e for compatibility reasons

hm	23. oct. 2008	REV 	2.0
	new code using _RMP_B

*)
          

METHOD SetRMP
  VAR_INPUT
    RMP : BYTE;
  END_VAR
                  THIS^.OUT:=RMP;
THIS^.rmp.SetRMP(RMP);
                
END_METHOD
END_FUNCTION_BLOCK

FUNCTION SwapWordsToReal : REAL
  VAR_INPUT
    wHi : WORD;
    wLo : WORD;
  END_VAR
  VAR
    dwVar : DWORD;
    pt_REAL : POINTER TO REAL;
  END_VAR

            dwVar := SHL(WORD_TO_DWORD(wHi),16) OR WORD_TO_DWORD(wLo);
pt_REAL := ADR(dwVar);
SwapWordsToReal := pt_REAL^;
          
END_FUNCTION

PROGRAM PLC_PRG_MAIN
  VAR
    MqttPushbuttonPrefix : STRING(100) := 'Devices/PLC/House/Out/DigitalInputs/Pushbuttons/';  (* INPUT FUNCTION BLOCKS *)
    FB_DI_PB_001 : FB_INPUT_PUSHBUTTON_MQTT;
    FB_DI_PB_002 : FB_INPUT_PUSHBUTTON_MQTT;
    FB_DI_PB_003 : FB_INPUT_PUSHBUTTON_MQTT;
    FB_DI_PB_004 : FB_INPUT_PUSHBUTTON_MQTT;
    FB_DI_PB_005 : FB_INPUT_PUSHBUTTON_MQTT;
    FB_DI_PB_006 : FB_INPUT_PUSHBUTTON_MQTT;
    FB_DI_PB_007 : FB_INPUT_PUSHBUTTON_MQTT;
    FB_DI_PB_008 : FB_INPUT_PUSHBUTTON_MQTT;
    FB_DI_PB_009 : FB_INPUT_PUSHBUTTON_DIMMER_MQTT;
    FB_DI_PB_010 : FB_INPUT_PUSHBUTTON_MQTT;
    FB_DI_PB_011 : FB_INPUT_PUSHBUTTON_MQTT;
    FB_DI_PB_012 : FB_INPUT_PUSHBUTTON_MQTT;
    FB_DI_PB_013 : FB_INPUT_PUSHBUTTON_MQTT;
    FB_DI_PB_014 : FB_INPUT_PUSHBUTTON_MQTT;
    FB_DI_PB_015 : FB_INPUT_PUSHBUTTON_MQTT;
    FB_DI_PB_016 : FB_INPUT_PUSHBUTTON_MQTT;
    FB_DI_PB_017 : FB_INPUT_PUSHBUTTON_MQTT;
    FB_DI_PB_018 : FB_INPUT_PUSHBUTTON_MQTT;
    FB_DI_PB_019 : FB_INPUT_PUSHBUTTON_MQTT;
    FB_DI_PB_020 : FB_INPUT_PUSHBUTTON_MQTT;
    FB_DI_PB_021 : FB_INPUT_PUSHBUTTON_MQTT;
    FB_DI_PB_022 : FB_INPUT_PUSHBUTTON_MQTT;
    FB_DI_PB_023 : FB_INPUT_PUSHBUTTON_MQTT;
    FB_DI_PB_024 : FB_INPUT_PUSHBUTTON_MQTT;
    FB_DI_PB_025 : FB_INPUT_PUSHBUTTON_MQTT;
    FB_DI_PB_026 : FB_INPUT_PUSHBUTTON_MQTT;
    FB_DI_PB_027 : FB_INPUT_PUSHBUTTON_MQTT;
    FB_DI_PB_028 : FB_INPUT_PUSHBUTTON_MQTT;
    FB_DI_PB_029 : FB_INPUT_PUSHBUTTON_MQTT;
    FB_DI_PB_030 : FB_INPUT_PUSHBUTTON_MQTT;
    FB_DI_PB_031 : FB_INPUT_PUSHBUTTON_MQTT;
    FB_DI_PB_032 : FB_INPUT_PUSHBUTTON_MQTT;
    FB_DI_PB_033 : FB_INPUT_PUSHBUTTON_MQTT;
    FB_DI_PB_034 : FB_INPUT_PUSHBUTTON_MQTT;
    FB_DI_PB_035 : FB_INPUT_PUSHBUTTON_MQTT;
    FB_DI_PB_036 : FB_INPUT_PUSHBUTTON_MQTT;
    FB_DI_PB_037 : FB_INPUT_PUSHBUTTON_MQTT;
    FB_DI_PB_038 : FB_INPUT_PUSHBUTTON_MQTT;
    FB_DI_PB_039 : FB_INPUT_PUSHBUTTON_MQTT;
    FB_DI_PB_040 : FB_INPUT_PUSHBUTTON_MQTT;
    FB_DI_PB_041 : FB_INPUT_PUSHBUTTON_MQTT;
    FB_DI_PB_042 : FB_INPUT_PUSHBUTTON_MQTT;
    FB_DI_PB_043 : FB_INPUT_PUSHBUTTON_MQTT;
    FB_DI_PB_044 : FB_INPUT_PUSHBUTTON_MQTT;
    FB_DI_PB_045 : FB_INPUT_PUSHBUTTON_MQTT;
    FB_DI_PB_046 : FB_INPUT_PUSHBUTTON_MQTT;
    FB_DI_PB_047 : FB_INPUT_PUSHBUTTON_MQTT;
    FB_DI_PB_048 : FB_INPUT_PUSHBUTTON_MQTT;
    MqttPubSwitchPrefix : STRING(100) := 'Devices/PLC/House/Out/DigitalOutputs/';  (* OUTPUT FUNCTION BLOCKS *)
    MqttSubSwitchPrefix : STRING(100) := 'Devices/PLC/House/In/DigitalOutputs/';
    FB_DO_SW_001 : FB_OUTPUT_SWITCH_MQTT;
    FB_DO_SW_002 : FB_OUTPUT_SWITCH_MQTT;
    FB_DO_SW_003 : FB_OUTPUT_SWITCH_MQTT;
    FB_DO_SW_004 : FB_OUTPUT_SWITCH_MQTT;
    FB_DO_SW_005 : FB_OUTPUT_SWITCH_MQTT;
    FB_DO_SW_006 : FB_OUTPUT_SWITCH_MQTT;
    FB_DO_SW_007 : FB_OUTPUT_SWITCH_MQTT;
    FB_DO_SW_008 : FB_OUTPUT_SWITCH_MQTT;
    FB_DO_SW_009 : FB_OUTPUT_SWITCH_MQTT;
    FB_DO_SW_010 : FB_OUTPUT_SWITCH_MQTT;
    FB_DO_SW_011 : FB_OUTPUT_SWITCH_MQTT;
    FB_DO_SW_012 : FB_OUTPUT_SWITCH_MQTT;
    FB_DO_SW_013 : FB_OUTPUT_SWITCH_MQTT;
    FB_DO_SW_014 : FB_OUTPUT_SWITCH_MQTT;
    FB_DO_SW_015 : FB_OUTPUT_SWITCH_MQTT;
    FB_DO_SW_016 : FB_OUTPUT_SWITCH_MQTT;
    FB_DO_SW_017 : FB_OUTPUT_SWITCH_MQTT;
    FB_DO_SW_018 : FB_OUTPUT_SWITCH_MQTT;
    FB_DO_SW_019 : FB_OUTPUT_SWITCH_MQTT;
    FB_DO_SW_020 : FB_OUTPUT_SWITCH_MQTT;
    FB_DO_SW_021 : FB_OUTPUT_SWITCH_MQTT;
    FB_DO_SW_022 : FB_OUTPUT_SWITCH_MQTT;
    FB_DO_SW_023 : FB_OUTPUT_SWITCH_MQTT;
    FB_DO_SW_024 : FB_OUTPUT_SWITCH_MQTT;
    FB_DO_SW_025 : FB_OUTPUT_SWITCH_MQTT;
    FB_DO_SW_026 : FB_OUTPUT_SWITCH_MQTT;
    FB_DO_SW_027 : FB_OUTPUT_SWITCH_MQTT;
    FB_DO_SW_028 : FB_OUTPUT_SWITCH_MQTT;
    FB_DO_SW_029 : FB_OUTPUT_SWITCH_MQTT;
    FB_DO_SW_030 : FB_OUTPUT_SWITCH_MQTT;
    FB_DO_SW_031 : FB_OUTPUT_SWITCH_MQTT;
    FB_DO_SW_032 : FB_OUTPUT_SWITCH_MQTT;
    FB_DO_BISTABLE_001 : FB_OUTPUT_BISTABLE_MQTT;
    MqttPubCoverPrefix : STRING(100) := 'Devices/PLC/House/Out/Covers/';  (* COVER FUNCTION BLOCKS *)
    MqttSubCoverPrefix : STRING(100) := 'Devices/PLC/House/In/Covers/';
    FB_DO_COVER_001 : FB_OUTPUT_COVER_MQTT;
    MqttPubDimmerPrefix : STRING(100) := 'Devices/PLC/House/Out/Dimmers/';  (* DIMMER FUNCTION BLOCKS *)
    MqttSubDimmerPrefix : STRING(100) := 'Devices/PLC/House/In/Dimmers/';
    FB_AO_DIMMER_001 : FB_OUTPUT_DIMMER_MQTT;
    TestOUT : WORD;
    MqttPubVirtualPrefix : STRING(100) := 'Devices/PLC/House/Out/Virtuals/';  (* VIRTUAL FUNCTION BLOCKS *)
    MqttSubVirtualPrefix : STRING(100) := 'Devices/PLC/House/In/Virtuals/';
    FB_VIRTUAL_INT_001 : FB_VIRTUAL_INT_MQTT;
    FB_VIRTUAL_BOOL_001 : FB_VIRTUAL_BOOL_MQTT;
    FB_VIRTUAL_STRING_001 : FB_VIRTUAL_STRING_MQTT;
    FB_VIRTUAL_REAL_001 : FB_VIRTUAL_REAL_MQTT;
  END_VAR

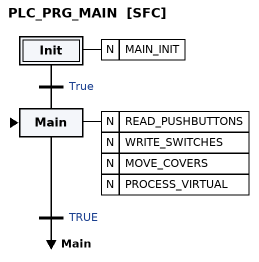
INITIAL_STEP Init:
  MAIN_INIT(N);
END_STEP
TRANSITION FROM Init TO Main
  := True;
END_TRANSITION
STEP Main:
  READ_PUSHBUTTONS(N);
  WRITE_SWITCHES(N);
  MOVE_COVERS(N);
  PROCESS_VIRTUAL(N);
END_STEP
TRANSITION FROM Main TO Main
  := TRUE;
END_TRANSITION

ACTION READ_PUSHBUTTONS:
                      FB_DI_PB_001(PB:= DI_001); (* Provide the input FB the correct phyical input to validate each cyclus *)
FB_DI_PB_002(PB:= DI_002);
FB_DI_PB_003(PB:= DI_003);
FB_DI_PB_004(PB:= DI_004);
FB_DI_PB_005(PB:= DI_005);
FB_DI_PB_006(PB:= DI_006);
FB_DI_PB_007(PB:= DI_007);
FB_DI_PB_008(PB:= DI_008);
FB_DI_PB_009(PB:= DI_009);
FB_DI_PB_010(PB:= DI_010);
FB_DI_PB_011(PB:= DI_011);
FB_DI_PB_012(PB:= DI_012);
FB_DI_PB_013(PB:= DI_013);
FB_DI_PB_014(PB:= DI_014);
FB_DI_PB_015(PB:= DI_015);
FB_DI_PB_016(PB:= DI_016);
FB_DI_PB_017(PB:= DI_017);
FB_DI_PB_018(PB:= DI_018);
FB_DI_PB_019(PB:= DI_019);
FB_DI_PB_020(PB:= DI_020);
FB_DI_PB_021(PB:= DI_021);
FB_DI_PB_022(PB:= DI_022);
FB_DI_PB_023(PB:= DI_023);
FB_DI_PB_024(PB:= DI_024);
FB_DI_PB_025(PB:= DI_025);
FB_DI_PB_026(PB:= DI_026);
FB_DI_PB_027(PB:= DI_027);
FB_DI_PB_028(PB:= DI_028);
FB_DI_PB_029(PB:= DI_029);
FB_DI_PB_030(PB:= DI_030);
FB_DI_PB_031(PB:= DI_031);
FB_DI_PB_032(PB:= DI_032);
FB_DI_PB_033(PB:= DI_033);
FB_DI_PB_034(PB:= DI_034);
FB_DI_PB_035(PB:= DI_035);
FB_DI_PB_036(PB:= DI_036);
FB_DI_PB_037(PB:= DI_037);
FB_DI_PB_038(PB:= DI_038);
FB_DI_PB_039(PB:= DI_039);
FB_DI_PB_040(PB:= DI_040);
FB_DI_PB_041(PB:= DI_041);
FB_DI_PB_042(PB:= DI_042);
FB_DI_PB_043(PB:= DI_043);
FB_DI_PB_044(PB:= DI_044);
FB_DI_PB_045(PB:= DI_045);
FB_DI_PB_046(PB:= DI_046);
FB_DI_PB_047(PB:= DI_047);
FB_DI_PB_048(PB:= DI_048);
                    
END_ACTION

ACTION WRITE_SWITCHES:
                      FB_DO_SW_001(OUT	=>		DO_001,										(* couple the function block to the physical output *)
	PRIO_HIGH				:=FALSE,  									(* brings the output high regardless of other input values *)
	PRIO_LOW				:=FALSE, 									(* brings the output low regardless of other input values. NOTE: PRIO_HIGH overrules PRIO_LOW input *)
	TOGGLE					:=FB_DI_PB_009.SINGLE 						(* for toggling the output *)	
);

FB_DO_SW_002(OUT => DO_002		,PRIO_HIGH:=FALSE			,PRIO_LOW:=FALSE				,TOGGLE:=FB_DI_PB_009.DOUBLE	);
FB_DO_SW_003(OUT => DO_003		,PRIO_HIGH:=FALSE			,PRIO_LOW:=FALSE				,TOGGLE:=FB_DI_PB_009.LONG		);
FB_DO_SW_004(OUT => DO_004		,PRIO_HIGH:=FALSE			,PRIO_LOW:=FALSE				,TOGGLE:=FB_DI_PB_009.LONG		);
FB_DO_SW_005(OUT => DO_005		,PRIO_HIGH:=FALSE			,PRIO_LOW:=FALSE				,TOGGLE:=FB_DI_PB_009.LONG		);
FB_DO_SW_006(OUT => DO_006		,PRIO_HIGH:=FALSE			,PRIO_LOW:=FALSE				,TOGGLE:=FB_DI_PB_009.LONG		);
FB_DO_SW_007(OUT => DO_007		,PRIO_HIGH:=FALSE			,PRIO_LOW:=FALSE				,TOGGLE:=FB_DI_PB_009.LONG		);
FB_DO_SW_008(OUT => DO_008		,PRIO_HIGH:=FALSE			,PRIO_LOW:=FALSE				,TOGGLE:=FB_DI_PB_009.LONG		);
FB_DO_SW_009(OUT => DO_009		,PRIO_HIGH:=FALSE			,PRIO_LOW:=FALSE				,TOGGLE:=FALSE				);
FB_DO_SW_010(OUT => DO_010		,PRIO_HIGH:=FALSE			,PRIO_LOW:=FALSE				,TOGGLE:=FALSE				);
FB_DO_SW_011(OUT => DO_011		,PRIO_HIGH:=FALSE			,PRIO_LOW:=FALSE				,TOGGLE:=FALSE				);
FB_DO_SW_012(OUT => DO_012		,PRIO_HIGH:=FALSE			,PRIO_LOW:=FALSE				,TOGGLE:=FALSE				);
FB_DO_SW_013(OUT => DO_013		,PRIO_HIGH:=FALSE			,PRIO_LOW:=FALSE				,TOGGLE:=FALSE				);
FB_DO_SW_014(OUT => DO_014		,PRIO_HIGH:=FALSE			,PRIO_LOW:=FALSE				,TOGGLE:=FALSE				);
FB_DO_SW_015(OUT => DO_015		,PRIO_HIGH:=FALSE			,PRIO_LOW:=FALSE				,TOGGLE:=FALSE				);
FB_DO_SW_016(OUT => DO_016		,PRIO_HIGH:=FALSE			,PRIO_LOW:=FALSE				,TOGGLE:=FALSE				);
FB_DO_SW_017(OUT => DO_017		,PRIO_HIGH:=FALSE			,PRIO_LOW:=FALSE				,TOGGLE:=FALSE				);
FB_DO_SW_018(OUT => DO_018		,PRIO_HIGH:=FALSE			,PRIO_LOW:=FALSE				,TOGGLE:=FALSE				);
FB_DO_SW_019(OUT => DO_019		,PRIO_HIGH:=FALSE			,PRIO_LOW:=FALSE				,TOGGLE:=FALSE				);
FB_DO_SW_020(OUT => DO_020		,PRIO_HIGH:=FALSE			,PRIO_LOW:=FALSE				,TOGGLE:=FALSE				);
FB_DO_SW_021(OUT => DO_021		,PRIO_HIGH:=FALSE			,PRIO_LOW:=FALSE				,TOGGLE:=FALSE				);
FB_DO_SW_022(OUT => DO_022		,PRIO_HIGH:=FALSE			,PRIO_LOW:=FALSE				,TOGGLE:=FALSE				);
FB_DO_SW_023(OUT => DO_023		,PRIO_HIGH:=FALSE			,PRIO_LOW:=FALSE				,TOGGLE:=FALSE				);
FB_DO_SW_024(OUT => DO_024		,PRIO_HIGH:=FALSE			,PRIO_LOW:=FALSE				,TOGGLE:=FALSE				);
FB_DO_SW_025(OUT => DO_025		,PRIO_HIGH:=FALSE			,PRIO_LOW:=FALSE				,TOGGLE:=FALSE				);
FB_DO_SW_026(OUT => DO_026		,PRIO_HIGH:=FALSE			,PRIO_LOW:=FALSE				,TOGGLE:=FALSE				);
FB_DO_SW_027(OUT => DO_027		,PRIO_HIGH:=FALSE			,PRIO_LOW:=FALSE				,TOGGLE:=FALSE				);
FB_DO_SW_028(OUT => DO_028		,PRIO_HIGH:=FALSE			,PRIO_LOW:=FALSE				,TOGGLE:=FALSE				);
FB_DO_SW_029(OUT => DO_029		,PRIO_HIGH:=FALSE			,PRIO_LOW:=FALSE				,TOGGLE:=FALSE				);
FB_DO_SW_030(OUT => DO_030		,PRIO_HIGH:=FALSE			,PRIO_LOW:=FALSE				,TOGGLE:=FALSE				);


FB_AO_DIMMER_001(
	SINGLE:=FB_DI_PB_041.SINGLE,
	LONG:=FB_DI_PB_041.LONG, 
	P_LONG:=FB_DI_PB_041.P_LONG, 
	Q_OUT => TestOUT,
	SET:=  FB_DI_PB_041.DOUBLE,
	VAL:=125
);

FB_DO_BISTABLE_001();
                    
END_ACTION

ACTION MAIN_INIT:
                      (* INIT DIGITAL INPUT STUFF *)
FB_DI_PB_001.InitMqtt(MQTTPublishPrefix:= ADR(MqttPushbuttonPrefix),	(* pointer to string prefix for the mqtt publish topic *)
	pMqttPublishQueue := ADR(MqttVariables.fbMqttPublishQueue)		(* pointer to MqttPublishQueue to send a new Mqtt event *)
);
FB_DI_PB_002.InitMqtt(MQTTPublishPrefix:= ADR(MqttPushbuttonPrefix),	pMqttPublishQueue := ADR(MqttVariables.fbMqttPublishQueue));
FB_DI_PB_003.InitMqtt(MQTTPublishPrefix:= ADR(MqttPushbuttonPrefix),	pMqttPublishQueue := ADR(MqttVariables.fbMqttPublishQueue));
FB_DI_PB_004.InitMqtt(MQTTPublishPrefix:= ADR(MqttPushbuttonPrefix),	pMqttPublishQueue := ADR(MqttVariables.fbMqttPublishQueue));
FB_DI_PB_005.InitMqtt(MQTTPublishPrefix:= ADR(MqttPushbuttonPrefix),	pMqttPublishQueue := ADR(MqttVariables.fbMqttPublishQueue));
FB_DI_PB_006.InitMqtt(MQTTPublishPrefix:= ADR(MqttPushbuttonPrefix),	pMqttPublishQueue := ADR(MqttVariables.fbMqttPublishQueue));
FB_DI_PB_007.InitMqtt(MQTTPublishPrefix:= ADR(MqttPushbuttonPrefix),	pMqttPublishQueue := ADR(MqttVariables.fbMqttPublishQueue));
FB_DI_PB_008.InitMqtt(MQTTPublishPrefix:= ADR(MqttPushbuttonPrefix),	pMqttPublishQueue := ADR(MqttVariables.fbMqttPublishQueue));
FB_DI_PB_009.InitMqtt(MQTTPublishPrefix:= ADR(MqttPushbuttonPrefix),	pMqttPublishQueue := ADR(MqttVariables.fbMqttPublishQueue), TRUE, MQTT.QoS.ExactlyOnce, 5);
FB_DI_PB_010.InitMqtt(MQTTPublishPrefix:= ADR(MqttPushbuttonPrefix),	pMqttPublishQueue := ADR(MqttVariables.fbMqttPublishQueue));
FB_DI_PB_011.InitMqtt(MQTTPublishPrefix:= ADR(MqttPushbuttonPrefix),	pMqttPublishQueue := ADR(MqttVariables.fbMqttPublishQueue));
FB_DI_PB_012.InitMqtt(MQTTPublishPrefix:= ADR(MqttPushbuttonPrefix),	pMqttPublishQueue := ADR(MqttVariables.fbMqttPublishQueue));
FB_DI_PB_013.InitMqtt(MQTTPublishPrefix:= ADR(MqttPushbuttonPrefix),	pMqttPublishQueue := ADR(MqttVariables.fbMqttPublishQueue));
FB_DI_PB_014.InitMqtt(MQTTPublishPrefix:= ADR(MqttPushbuttonPrefix),	pMqttPublishQueue := ADR(MqttVariables.fbMqttPublishQueue));
FB_DI_PB_015.InitMqtt(MQTTPublishPrefix:= ADR(MqttPushbuttonPrefix),	pMqttPublishQueue := ADR(MqttVariables.fbMqttPublishQueue));
FB_DI_PB_016.InitMqtt(MQTTPublishPrefix:= ADR(MqttPushbuttonPrefix),	pMqttPublishQueue := ADR(MqttVariables.fbMqttPublishQueue));
FB_DI_PB_041.InitMqtt(MQTTPublishPrefix:= ADR(MqttPushbuttonPrefix),	pMqttPublishQueue := ADR(MqttVariables.fbMqttPublishQueue));

(* INIT DIMMER OUTPUT STUFF *)
FB_AO_DIMMER_001.InitMQTT(MQTTPublishPrefix:= ADR(MqttPubDimmerPrefix),    (* pointer to string prefix for the MQTT publish topic *)
	MQTTSubscribePrefix:= ADR(MqttSubDimmerPrefix),							(* pointer to string prefix for the MQTT subscribe topic *)
    pMQTTPublishQueue := ADR(MQTTVariables.fbMQTTPublishQueue),         (* pointer to MQTTPublishQueue to send a new MQTT event *)
	pMqttCallbackCollector := ADR(MqttVariables.collector_FB_DIMMER_MQTT),	(* pointer to CallbackCollector to receive Mqtt subscription events *)
    TRUE,                                                               (* specify whether dimmer value should be outputted on MQTT topic *)
    MQTT.QoS.ExactlyOnce,                                            (* specify the QoS for the dimmer mqtt events (values 0-255) *)    
    5                                                                   (* specify the resolution for the dimmer mqtt events *)     
);

(* ALTER THE DIMMER OUTPUT DEFAULT BEHAVIOR *)
FB_AO_DIMMER_001.ConfigureFunctionBlock(
	T_Debounce:=T#10MS,
	T_Reconfig:=T#10S,
	T_On_Max:=T#0S,
	T_Dimm_Start:=T#400MS,
	T_Dimm:=T#3S,
	Min_On:=50,
	Max_On:=255,
	Soft_Dimm:=TRUE,
	Rst_Out:=FALSE,
	OUT_LinearScaleMin:=11000,
	OUT_LinearScaleMax:=32767
);


